ACTION AxisModules:
//*******************************************************************************************************************
// Moduli asse (Core: FB_AxisModule): ingressi dalla macchina, chiamate, uscite verso Safety e allarmi
//*******************************************************************************************************************
// In uso: per un asse aggiunto vale la presenza nei parametri macchina (Hmi.Param); per i sei assi storici le
// regole di prima. UR2 e UR_SIM: e' in uso uno solo dei due (ur2InUse); prima un'unica istanza di jog e di reset cambiava asse.
FOR i := 1 TO Mach.MAX_AXIS_CFG DO
	axisInUse[i] := Mach.aAxisCfg[i].bDefined AND Hmi.Param.aAxis[i].bPresent;
END_FOR
axisInUse[Mach.AX_USEL]		:= TRUE;
axisInUse[Mach.AX_USER]		:= TRUE;
axisInUse[Mach.AX_ERL]		:= TRUE;
axisInUse[Mach.AX_ERR]		:= TRUE;
axisInUse[Mach.AX_UR2]		:= ur2InUse;
axisInUse[Mach.AX_UR_SIM]	:= NOT ur2InUse;

// Ingressi comuni, dalla configurazione dell'asse (FB_MachineConfig)
mpgSelector := DINT_TO_UINT(stMpgEncoder.diSelector1);
FOR i := 1 TO Mach.MAX_AXIS_CFG DO
	IF Mach.aAxisCfg[i].bDefined THEN
		aAxisMod[i].bPowerEnable		:= axisInUse[i] AND motorsOn AND Safety.EmergenzaResettata;
		aAxisMod[i].fOverride			:= axisOverride;
		aAxisMod[i].bUseSoEReset		:= Mach.aAxisCfg[i].bSoEReset;
		aAxisMod[i].bSoEResetRequest	:= Safety.PulsanteResetEmergenza;
		aAxisMod[i].tPoweredOffDelay	:= tMotorsOffDelay;
		aAxisMod[i].bResetExecute		:= resetAxesCmd AND axisInUse[i];
		// Jog dal volantino: solo in manuale e con il ciclo fermo, l'asse scelto dal selettore.
		jogSelected := manualMode AND state = E_CycleState.Idle AND axisInUse[i]
			AND NOT calibStart[i] AND aAxisMod[i].nCalibrationStep = 0
			AND Mach.aAxisCfg[i].nMpgSelector <> 0 AND Mach.aAxisCfg[i].nMpgSelector = mpgSelector
			AND stMpgEncoder.diSafetySwitch;
		// Jog dall'HMI (stesse condizioni; i motori in manuale li tiene accesi il consenso del volantino).
		jogHmi := hmiConnected AND manualMode AND state = E_CycleState.Idle AND axisInUse[i] AND Hmi.Live.nJogAxis = i
			AND NOT calibStart[i] AND aAxisMod[i].nCalibrationStep = 0;
		aAxisMod[i].bJogForward			:= (jogSelected AND stMpgEncoder.eDirection = MC_Direction.MC_Positive_Direction)
			OR (jogHmi AND Hmi.Live.nJogDirection > 0);
		aAxisMod[i].bJogBackward		:= (jogSelected AND stMpgEncoder.eDirection = MC_Direction.MC_Negative_Direction)
			OR (jogHmi AND Hmi.Live.nJogDirection < 0);
		aAxisMod[i].fJogVelocity		:= Mach.aAxisCfg[i].fJogVelocity;
		aAxisMod[i].fJogAcceleration	:= Mach.aAxisCfg[i].fJogAcceleration;
		aAxisMod[i].fJogDeceleration	:= Mach.aAxisCfg[i].fJogDeceleration;
		aAxisMod[i].fJogJerk			:= Mach.aAxisCfg[i].fJogJerk;
		aAxisMod[i].bCalibrationStart	:= calibStart[i];
		aAxisMod[i].bUseCalibrationPos	:= calibUsePos[i];
		aAxisMod[i].fCalibrationPos		:= calibPos[i];
		aAxisMod[i].bWriteLimits		:= (i = limitsKickAxis);	// un asse alla volta (vedi fine AxisModules)
		// Limiti di un asse aggiunto dai parametri HMI; per gli assi storici li sovrascrive il blocco sotto.
		aAxisMod[i].fUpperLimit			:= Hmi.Param.aAxis[i].fUpperLimit;
		aAxisMod[i].fLowerLimit			:= Hmi.Param.aAxis[i].fLowerLimit;
	END_IF
END_FOR

// Calibrazione: comando e quota da HmiInputs (comando Calibrate), quota standard (GVL Calibration), datum di sicurezza
aAxisMod[Mach.AX_ERL].fHomePosition			:= Calibration.ERLHomePosition;
aAxisMod[Mach.AX_ERL].bDatumRequest			:= Safety.ERLDatumRequest;
aAxisMod[Mach.AX_ERL].bDatumDone			:= Safety.ERLDatumDone;

aAxisMod[Mach.AX_USEL].fHomePosition		:= Calibration.USELHomePosition;
aAxisMod[Mach.AX_USEL].bDatumRequest		:= Safety.USELDatumRquest;
aAxisMod[Mach.AX_USEL].bDatumDone			:= Safety.USELDatumDone;

aAxisMod[Mach.AX_UR2].fHomePosition			:= Calibration.URHomePosition;
aAxisMod[Mach.AX_UR2].bDatumRequest			:= Safety.URDatumRequest;
aAxisMod[Mach.AX_UR2].bDatumDone			:= Safety.URDatumDone;

aAxisMod[Mach.AX_ERR].fHomePosition			:= Calibration.ERRHomePosition;
aAxisMod[Mach.AX_ERR].bDatumRequest			:= Safety.ERRDatumRequest;
aAxisMod[Mach.AX_ERR].bDatumDone			:= Safety.ERRDatumDone;

aAxisMod[Mach.AX_USER].fHomePosition		:= Calibration.USERHomePosition;
aAxisMod[Mach.AX_USER].bDatumRequest		:= Safety.USERDatumRequest;
aAxisMod[Mach.AX_USER].bDatumDone			:= Safety.USERDatumDone;

// Limiti software dai parametri macchina (copia locale parametersRx). Il minimo delle USE non scende sotto
// il finecorsa della morsa montata (urUSE*MinPosition senza UR2, ur2USE*MinPosition con UR2).
aAxisMod[Mach.AX_ERL].fUpperLimit	:= parametersRx.ErLUpperLimit;
aAxisMod[Mach.AX_ERL].fLowerLimit	:= parametersRx.ErLLowerLimit;
aAxisMod[Mach.AX_USEL].fUpperLimit	:= parametersRx.UseLUpperLimit;
aAxisMod[Mach.AX_USEL].fLowerLimit	:= MAX(parametersRx.UseLLowerLimit, SEL(ur2InUse, urUSELMinPosition, ur2USELMinPosition));
aAxisMod[Mach.AX_UR2].fUpperLimit	:= parametersRx.UrRUpperLimit;
aAxisMod[Mach.AX_UR2].fLowerLimit	:= parametersRx.UrRLowerLimit;
aAxisMod[Mach.AX_ERR].fUpperLimit	:= parametersRx.ErRUpperLimit;
aAxisMod[Mach.AX_ERR].fLowerLimit	:= parametersRx.ErRLowerLimit;
aAxisMod[Mach.AX_USER].fUpperLimit	:= parametersRx.UseRUpperLimit;
aAxisMod[Mach.AX_USER].fLowerLimit	:= MAX(parametersRx.UseRLowerLimit, SEL(ur2InUse, urUSERMinPosition, ur2USERMinPosition));

// Chiamate (un asse NC per modulo)
aAxisMod[Mach.AX_USEL](stAxis := USEL);
aAxisMod[Mach.AX_USER](stAxis := USER);
aAxisMod[Mach.AX_ERL](stAxis := ERL);
aAxisMod[Mach.AX_ERR](stAxis := ERR);
aAxisMod[Mach.AX_UR2](stAxis := UR2);
aAxisMod[Mach.AX_UR_SIM](stAxis := UR_SIM);

// Uscite verso la sicurezza (lo stato della calibrazione per l'HMI e' in HmiOutputs)
// ERLDatumExecute non si azzera mai, come prima (la riga in InitCyclic era commentata): da verificare sullo schema safety.
IF aAxisMod[Mach.AX_ERL].bDatumExecute THEN
	Safety.ERLDatumExecute := TRUE;
END_IF
Safety.USELDatumExecute		:= aAxisMod[Mach.AX_USEL].bDatumExecute;
Safety.URDatumExecute		:= aAxisMod[Mach.AX_UR2].bDatumExecute;
Safety.ERRDatumExecute		:= aAxisMod[Mach.AX_ERR].bDatumExecute;
Safety.USERDatumExecute		:= aAxisMod[Mach.AX_USER].bDatumExecute;

// Esiti per la macchina a stati (letti nel ciclo dopo, come prima) e allarmi chiesti dai moduli
axesResetDone := TRUE;
axesResetError := FALSE;
axesResetErrorId := 0;
limitsBusy := FALSE;
FOR i := 1 TO Mach.MAX_AXIS_CFG DO
	IF Mach.aAxisCfg[i].bDefined THEN
		IF axisInUse[i] THEN
			axesResetDone := axesResetDone AND aAxisMod[i].bResetDone;
			IF aAxisMod[i].bResetError THEN
				axesResetError := TRUE;
				axesResetErrorId := MAX(axesResetErrorId, aAxisMod[i].nResetErrorId);
			END_IF
		END_IF
		limitsBusy := limitsBusy OR aAxisMod[i].bLimitsBusy;
		limitsFailed := limitsFailed OR aAxisMod[i].bLimitsError;
		CASE aAxisMod[i].eAlarm OF
			E_AxisAlarm.Calibration:
				RaiseAlarm(Id := Mach.aAxisCfg[i].nCalibrationAlarmId, Info := aAxisMod[i].nAlarmInfo);
			E_AxisAlarm.Limits:
				RaiseAlarm(Id := Mach.aAxisCfg[i].nLimitsAlarmId, Info := aAxisMod[i].nAlarmInfo);
		END_CASE
	END_IF
END_FOR

// Scrittura dei limiti un asse alla volta, come il vecchio ParameterWriteManager (MC_WriteParameter, non
// persistente: vedi FB_AxisModule). Un asse che fallisce non ferma i successivi.
// Fine: l'HMI aspetta Hmi.Sts.bWriteParametersDone FALSE -> TRUE (resta FALSE se un asse fallisce).
limitsKickAxis := 0;
IF limitsWriting AND NOT limitsBusy THEN
	FOR i := limitsAxis + 1 TO Mach.MAX_AXIS_CFG DO
		// asse simulato: nessun limite da scrivere
		IF limitsKickAxis = 0 AND Mach.aAxisCfg[i].bDefined AND i <> Mach.AX_UR_SIM THEN
			limitsKickAxis := i;
		END_IF
	END_FOR
	IF limitsKickAxis <> 0 THEN
		limitsAxis := limitsKickAxis;
	ELSE
		limitsWriting := FALSE;
		writeParametersDone := NOT limitsFailed;
	END_IF
END_IF
END_ACTION

ACTION DiagUpdate:
// Stato dei canali e storico dei cambi di passo nella GVL Diag (letta dall'HMI in un blocco).
FOR i := 0 TO 2 DO
	IF state = E_CycleState.HomingRun OR state = E_CycleState.HomingPrepare THEN
		Diag.Data.aChannel[i].bUsed := ProgramDB.homing.task[i].active;
	ELSE
		Diag.Data.aChannel[i].bUsed := ProgramDB.sequence[seqIdx].task[i].active;
	END_IF
	Diag.Data.aChannel[i].bDone := channelDone[i];
	Diag.Data.aChannel[i].bMWaiting := in_stNciToPlc[i].HskMFuncReq = 1 AND out_stPlcToNci[i].MFuncGranted = 0;
	IF in_stNciToPlc[i].HskMFuncReq = 1 THEN
		Diag.Data.aChannel[i].nMFunc := in_stNciToPlc[i].HskMFuncNo;
	ELSE
		Diag.Data.aChannel[i].nMFunc := 0;
	END_IF
	fbMFuncWait[i](IN := Diag.Data.aChannel[i].bMWaiting, PT := T#24H);
	Diag.Data.aChannel[i].tMWait := fbMFuncWait[i].ET;
	Diag.Data.aChannel[i].nItpState := udiItpState[i];
END_FOR
Diag.Data.aChannel[0].nLineNo := lineNo1;
Diag.Data.aChannel[1].nLineNo := lineNo2;
Diag.Data.aChannel[2].nLineNo := lineNo3;

// Sequenze attive: si ricontano solo quando arriva un programma nuovo (e al primo giro).
IF newProgramTrigger OR NOT diagSeqCounted THEN
	diagSeqCounted := TRUE;
	diagSeqIdx := 0;
	WHILE diagSeqIdx < Size.MAX_SEQUENCE AND_THEN ProgramDB.sequence[diagSeqIdx].active DO
		diagSeqIdx := diagSeqIdx + 1;
	END_WHILE
	Diag.Data.nSeqCount := diagSeqIdx;
END_IF

Diag.Data.eCycleEndReason := cycleEndReason;
IF state = E_CycleState.Centering THEN
	Diag.Data.nSubStep := fbCentering.nStep;
ELSE
	Diag.Data.nSubStep := fbSeq.eStep;
END_IF

fbDiagLog(
	nState		:= state,
	nSeqIdx		:= seqIdx,
	nAbortState	:= E_CycleState.Abort,
	nAlarmCount	:= Alarms.RaisedCount,
	nAlarmId	:= Alarms.LastRaisedId,
	nAlarmInfo	:= Alarms.LastRaisedInfo,
	stDiag		:= Diag.Data);
END_ACTION

ACTION DriveStatusManager:
// Calcola stato drive e consenso motori per HMI.
allDrivesEnabled := (bMotorsOnStatus[0] OR NOT Machine.parametersRx.USELPresent) AND 
					(bMotorsOnStatus[1] OR NOT Machine.parametersRx.ERLPresent) AND 
					(bMotorsOnStatus[2] OR NOT ur2InUse) AND 
					(bMotorsOnStatus[3] OR NOT Machine.parametersRx.USERPresent) AND
					(bMotorsOnStatus[4] OR NOT Machine.parametersRx.ERRPresent);
					
drivesError := (USEL.NcToPlc.ErrorCode <> 0 AND Machine.parametersRx.USELPresent) OR
			   (ERL.NcToPlc.ErrorCode <> 0 AND Machine.parametersRx.ERLPresent) OR
			   (USER.NcToPlc.ErrorCode <> 0 AND Machine.parametersRx.USERPresent) OR
			   (ERR.NcToPlc.ErrorCode <> 0 AND Machine.parametersRx.ERRPresent) OR
			   (UR2.NcToPlc.ErrorCode <> 0 AND ur2InUse);

//fbMotorsOffTrigger(CLK := allDrivesEnabled, Q => motorsOffTrigger);
fbSelectorOffTrigger(CLK := Safety.ModoAuto1Op, Q=> autoModeTrigger);

IF drivesError OR  motorsOffTrigger THEN
	motorsOn := FALSE;
END_IF
END_ACTION

ACTION HmiInputs:
//*******************************************************************************************************************
// Ingressi dall'HMI (GVL Hmi, contratto in docs/ADS_CONTRACT_V2.md) nelle variabili interne
//*******************************************************************************************************************
fbHmiWatchdog(nCounter := Hmi.Live.nWatchdog);
hmiConnected := fbHmiWatchdog.bAlive;

// Comandi con numero di sequenza: valgono un ciclo.
hmiStartCmd := FALSE;
hmiStopCmd := FALSE;
hmiResetCmd := FALSE;
hmiMotorsOnCmd := FALSE;
hmiMotorsOffCmd := FALSE;
hmiProgramLoadedCmd := FALSE;
hmiWriteParamsCmd := FALSE;
FOR i := 1 TO Mach.MAX_AXIS_CFG DO
	calibStart[i] := FALSE;
END_FOR

fbHmiCmd(stCmd := Hmi.Cmd);
IF fbHmiCmd.bNew THEN
	CASE Hmi.Cmd.eCommand OF
		E_HmiCommand.Start:
			hmiStartCmd := TRUE;
			fbHmiCmd.Ack(E_HmiResult.Accepted);
		E_HmiCommand.Stop:
			hmiStopCmd := TRUE;
			fbHmiCmd.Ack(E_HmiResult.Accepted);
		E_HmiCommand.Reset:
			hmiResetCmd := TRUE;
			fbHmiCmd.Ack(E_HmiResult.Accepted);
		E_HmiCommand.MotorsOn:
			hmiMotorsOnCmd := TRUE;
			fbHmiCmd.Ack(E_HmiResult.Accepted);
		E_HmiCommand.MotorsOff:
			hmiMotorsOffCmd := TRUE;
			fbHmiCmd.Ack(E_HmiResult.Accepted);
		E_HmiCommand.ProgramLoaded:
			hmiProgramLoadedCmd := TRUE;
			fbHmiCmd.Ack(E_HmiResult.Accepted);
		E_HmiCommand.WriteParameters:
			// Parametri macchina dell'HMI -> struttura persistente usata da tutto il PLC (Machine.parametersRx).
			Machine.parametersRx.EnableSirenOverride	:= Hmi.Param.bEnableSirenOverride;
			Machine.parametersRx.ERLPresent			:= Hmi.Param.aAxis[Mach.AX_ERL].bPresent;
			Machine.parametersRx.ERLCalibrated		:= Hmi.Param.aAxis[Mach.AX_ERL].bCalibrated;
			Machine.parametersRx.ERLCheckDone		:= Hmi.Param.aAxis[Mach.AX_ERL].bCheckDone;
			Machine.parametersRx.ErLUpperLimit		:= Hmi.Param.aAxis[Mach.AX_ERL].fUpperLimit;
			Machine.parametersRx.ErLLowerLimit		:= Hmi.Param.aAxis[Mach.AX_ERL].fLowerLimit;
			Machine.parametersRx.USELPresent		:= Hmi.Param.aAxis[Mach.AX_USEL].bPresent;
			Machine.parametersRx.USELCalibrated		:= Hmi.Param.aAxis[Mach.AX_USEL].bCalibrated;
			Machine.parametersRx.USELCheckDone		:= Hmi.Param.aAxis[Mach.AX_USEL].bCheckDone;
			Machine.parametersRx.UseLUpperLimit		:= Hmi.Param.aAxis[Mach.AX_USEL].fUpperLimit;
			Machine.parametersRx.UseLLowerLimit		:= Hmi.Param.aAxis[Mach.AX_USEL].fLowerLimit;
			Machine.parametersRx.UR2Present			:= Hmi.Param.aAxis[Mach.AX_UR2].bPresent;
			Machine.parametersRx.UR2Calibrated		:= Hmi.Param.aAxis[Mach.AX_UR2].bCalibrated;
			Machine.parametersRx.ER2CheckDone		:= Hmi.Param.aAxis[Mach.AX_UR2].bCheckDone;
			Machine.parametersRx.UrRUpperLimit		:= Hmi.Param.aAxis[Mach.AX_UR2].fUpperLimit;
			Machine.parametersRx.UrRLowerLimit		:= Hmi.Param.aAxis[Mach.AX_UR2].fLowerLimit;
			Machine.parametersRx.ERRPresent			:= Hmi.Param.aAxis[Mach.AX_ERR].bPresent;
			Machine.parametersRx.ERRCalibrated		:= Hmi.Param.aAxis[Mach.AX_ERR].bCalibrated;
			Machine.parametersRx.ERRCheckDone		:= Hmi.Param.aAxis[Mach.AX_ERR].bCheckDone;
			Machine.parametersRx.ErRUpperLimit		:= Hmi.Param.aAxis[Mach.AX_ERR].fUpperLimit;
			Machine.parametersRx.ErRLowerLimit		:= Hmi.Param.aAxis[Mach.AX_ERR].fLowerLimit;
			Machine.parametersRx.USERPresent		:= Hmi.Param.aAxis[Mach.AX_USER].bPresent;
			Machine.parametersRx.USERCalibrated		:= Hmi.Param.aAxis[Mach.AX_USER].bCalibrated;
			Machine.parametersRx.USERCheckDone		:= Hmi.Param.aAxis[Mach.AX_USER].bCheckDone;
			Machine.parametersRx.UseRUpperLimit		:= Hmi.Param.aAxis[Mach.AX_USER].fUpperLimit;
			Machine.parametersRx.UseRLowerLimit		:= Hmi.Param.aAxis[Mach.AX_USER].fLowerLimit;
			hmiWriteParamsCmd := TRUE;
			fbHmiCmd.Ack(E_HmiResult.Accepted);
		E_HmiCommand.Calibrate:
			IF Hmi.Cmd.nAxis < 1 OR Hmi.Cmd.nAxis > Mach.MAX_AXIS_CFG THEN
				fbHmiCmd.Ack(E_HmiResult.InvalidArgument);
			ELSIF NOT Mach.aAxisCfg[Hmi.Cmd.nAxis].bDefined OR Mach.aAxisCfg[Hmi.Cmd.nAxis].nCalibrationAlarmId = 0 THEN
				fbHmiCmd.Ack(E_HmiResult.InvalidArgument);		// asse senza calibrazione (es. UR_SIM)
			ELSIF NOT manualMode OR NOT Safety.ModoManuale OR state <> E_CycleState.Idle
				OR limitsWriting OR limitsRequest OR limitsStart OR aAxisMod[Hmi.Cmd.nAxis].bLimitsBusy THEN
				fbHmiCmd.Ack(E_HmiResult.Rejected);		// solo da fermo in manuale, senza scritture limiti
			ELSIF aAxisMod[Hmi.Cmd.nAxis].nCalibrationStep <> 0 THEN
				fbHmiCmd.Ack(E_HmiResult.Rejected);				// calibrazione gia' in corso
			ELSE
				calibStart[Hmi.Cmd.nAxis] := TRUE;
				calibUsePos[Hmi.Cmd.nAxis] := Hmi.Cmd.bFlag;
				calibPos[Hmi.Cmd.nAxis] := Hmi.Cmd.fValue;
				fbHmiCmd.Ack(E_HmiResult.Accepted);
			END_IF
		E_HmiCommand.SetCount:
			IF Hmi.Cmd.nValue >= 0 AND Hmi.Cmd.nValue <= 65535 THEN
				count := DINT_TO_UINT(Hmi.Cmd.nValue);
				fbHmiCmd.Ack(E_HmiResult.Accepted);
			ELSE
				fbHmiCmd.Ack(E_HmiResult.InvalidArgument);
			END_IF
	ELSE
		fbHmiCmd.Ack(E_HmiResult.UnknownCommand);
	END_CASE
END_IF

// Valori continui (Hmi.Live). Con l'HMI scollegata restano gli ultimi scritti, tranne il test uscite che si spegne.
hmiOverride := Hmi.Live.fOverride;
autoLoopMode := Hmi.Live.bLoopMode;
ncSingleBlock := Hmi.Live.nNcMode = 1;
hmiForce := hmiConnected AND Hmi.Live.bForceOutputs;
FOR i := 1 TO Mach.MAX_VALVE DO
	valveForce[i] := Hmi.Live.aValveForce[i];
END_FOR

// Pulsanti
hmiStop := hmiStopCmd;
hmiReset := hmiResetCmd;
END_ACTION

ACTION HmiOutputs:
//*******************************************************************************************************************
// Stato per l'HMI (GVL Hmi): configurazione e stato, un blocco ciascuno
//*******************************************************************************************************************
Hmi.Cfg.nInterfaceVersion	:= 2;
Hmi.Cfg.sMachine			:= 'Aut260045';
Hmi.Cfg.nMaxSequence		:= Size.MAX_SEQUENCE;
Hmi.Cfg.nMaxTask			:= Size.MAX_TASK;
Hmi.Cfg.nMaxAction			:= Size.MAX_ACTION;
Hmi.Cfg.nMaxPosition		:= Size.MAX_POSITION;
Hmi.Cfg.nMaxMacro			:= Size.MAX_MACRO;
Hmi.Cfg.nMaxAxisInGroup		:= Size.MAX_AXIS;
Hmi.Cfg.nChannels			:= Core_Param.MAX_CHANNEL;

FOR i := 1 TO Mach.MAX_AXIS_CFG DO
	Hmi.Cfg.aAxis[i].bDefined	:= Mach.aAxisCfg[i].bDefined;
	Hmi.Cfg.aAxis[i].sName		:= Mach.aAxisCfg[i].sName;
	Hmi.Cfg.aAxis[i].nOption	:= Mach.aAxisCfg[i].nMpgSelector;
	Hmi.Sts.aAxis[i].fActPos			:= Mach.aAxisCfg[i].fActPos;
	Hmi.Sts.aAxis[i].fActVelo			:= Mach.aAxisCfg[i].fActVelo;
	Hmi.Sts.aAxis[i].nErrorCode			:= Mach.aAxisCfg[i].nErrorCode;
	Hmi.Sts.aAxis[i].bEnabled			:= Mach.aAxisCfg[i].bDefined AND NOT Mach.aAxisCfg[i].bDisabled;
	Hmi.Sts.aAxis[i].bMoving			:= Mach.aAxisCfg[i].bMoving;
	Hmi.Sts.aAxis[i].bInUse				:= axisInUse[i];
	Hmi.Sts.aAxis[i].nCalibrationStep	:= aAxisMod[i].nCalibrationStep;
	Hmi.Sts.aAxis[i].bCalibrated		:= aAxisMod[i].bCalibrated;
	Hmi.Sts.aAxis[i].bLimitsBusy		:= aAxisMod[i].bLimitsBusy;
END_FOR
Hmi.Sts.aAxis[Mach.AX_ERL].fLastKnownPos	:= Machine.parametersTx.lastERLKnownPosition;
Hmi.Sts.aAxis[Mach.AX_USEL].fLastKnownPos	:= Machine.parametersTx.lastUSELKnownPosition;
Hmi.Sts.aAxis[Mach.AX_UR2].fLastKnownPos	:= Machine.parametersTx.lastUR2KnownPosition;
Hmi.Sts.aAxis[Mach.AX_ERR].fLastKnownPos	:= Machine.parametersTx.lastERRKnownPosition;
Hmi.Sts.aAxis[Mach.AX_USER].fLastKnownPos	:= Machine.parametersTx.lastUSERKnownPosition;

FOR i := 1 TO Mach.MAX_VALVE DO
	Hmi.Cfg.aValve[i].bDefined	:= Mach.aValve[i].pSet <> 0;
	Hmi.Cfg.aValve[i].sName		:= Mach.aValve[i].sName;
	Hmi.Cfg.aValve[i].nOption	:= SEL(Mach.aValve[i].eType = OUTPUT_ENUM.BISTABLE, 0, 1);
	IF Mach.aValve[i].pSet <> 0 THEN
		Hmi.Sts.aValve[i].bSet := Mach.aValve[i].pSet^;
	END_IF
	IF Mach.aValve[i].pReset <> 0 THEN
		Hmi.Sts.aValve[i].bReset := Mach.aValve[i].pReset^;
	END_IF
	IF Mach.aValve[i].pFbSet <> 0 THEN
		Hmi.Sts.aValve[i].bFbSet := Mach.aValve[i].pFbSet^;
	END_IF
	IF Mach.aValve[i].pFbReset <> 0 THEN
		Hmi.Sts.aValve[i].bFbReset := Mach.aValve[i].pFbReset^;
	END_IF
END_FOR

FOR i := 1 TO Core_Param.MAX_INPUT DO
	Hmi.Cfg.aInput[i].bDefined	:= Mach.aInput[i].pInput <> 0;
	Hmi.Cfg.aInput[i].sName		:= Mach.aInput[i].sName;
	IF Mach.aInput[i].pInput <> 0 THEN
		Hmi.Sts.aInput[i] := Mach.aInput[i].pInput^;
	END_IF
END_FOR

Hmi.Sts.nCmdAck				:= fbHmiCmd.nAck;
Hmi.Sts.eCmdResult			:= fbHmiCmd.eResult;
Hmi.Sts.bConnected			:= hmiConnected;
Hmi.Sts.nState				:= state;
Hmi.Sts.nSubStep			:= Diag.Data.nSubStep;
Hmi.Sts.eCycleEndReason		:= cycleEndReason;
Hmi.Sts.bIdle				:= programIdle;
Hmi.Sts.bCanExecute			:= programCanExecute;
Hmi.Sts.bRunning			:= programRunning;
Hmi.Sts.bStopped			:= programStopped;
Hmi.Sts.bAborted			:= programAborted;
Hmi.Sts.bHomingDone			:= homingDone;
Hmi.Sts.bManualMode			:= manualMode;
Hmi.Sts.bAutoMode			:= autoMode;
Hmi.Sts.bMotorsOn			:= allDrivesEnabled;
Hmi.Sts.bMotorsEnable		:= NOT drivesError;
Hmi.Sts.bLimitsWriting		:= limitsWriting;
Hmi.Sts.bWriteParametersDone := writeParametersDone;
Hmi.Sts.nCount				:= count;
Hmi.Sts.nSeqIdx				:= seqIdx;
Hmi.Sts.sProgramName		:= ProgramDB.parameters.prgName;
Hmi.Sts.aLineNo[0]			:= lineNo1;
Hmi.Sts.aLineNo[1]			:= lineNo2;
Hmi.Sts.aLineNo[2]			:= lineNo3;
FOR i := 0 TO 2 DO
	Hmi.Sts.aChannelDone[i] := channelDone[i];
END_FOR
Hmi.Sts.nMpgSelector		:= stMpgEncoder.diSelector1;
Hmi.Sts.nMpgSpeed			:= stMpgEncoder.diSelector2;
Hmi.Sts.aAlarmActive		:= Alarms.Active;
Hmi.Sts.aAlarmInfo			:= Alarms.Info;
END_ACTION

ACTION InitCyclic:
(*initialize data cyclic (every scan)*)
//*******************************************************************************************************************
// set FB defaults
//*******************************************************************************************************************
allDrivesEnabled	:= FALSE;
drivesError 		:= FALSE;


//Read Status
USEL.ReadStatus();
ERL.ReadStatus();
UR2.ReadStatus();
USER.ReadStatus();
ERR.ReadStatus();

resetAxesCmd								:= FALSE;	// FB_AxisModule: reset MC degli assi (passi 800 e 920)












fbMPGReadStatus.tUpdateTimerPt				:= T#5MS;
fbMPGReadStatus.uiScalingFactorDenominator	:= 300;
fbMPGReadStatus.uiScalingFactorNumerator	:= 1;
fbMpgReadStatus.uismoothingPercentage		:= 10;





parametersRx.ERLCalibrated					:= FALSE;
parametersRx.ERLPresent						:= FALSE;
parametersRx.ERRCalibrated					:= FALSE;
parametersRx.ERRPresent						:= FALSE;
parametersRx.UR2Calibrated					:= FALSE;
parametersRx.UR2Present						:= FALSE;
parametersRx.USELCalibrated					:= FALSE;
parametersRx.USELPresent					:= FALSE;
parametersRx.USERCalibrated					:= FALSE;
parametersRx.USERPresent					:= FALSE;
parametersRx.ERLCheckDone					:= FALSE;
parametersRx.USELCheckDone					:= FALSE;
parametersRx.ER2CheckDone					:= FALSE;
parametersRx.ERRCheckDone					:= FALSE;
parametersRx.USERCheckDone					:= FALSE;

fbCloseClampAfterCentering.IN				:= FALSE;
fbCloseClampAfterCentering.PT				:= T#1000MS;

waitForMove.IN 								:= FALSE;
waitForMove.PT 								:= T#1S;

startCondition								:= FALSE;
safeOverride								:= FALSE;
END_ACTION

ACTION InitOnce:
firstScan := FALSE;
END_ACTION

ACTION InputMapping:
//*******************************************************************************************************************
// Override, eventi dei comandi HMI, morsa in uso
//*******************************************************************************************************************
axisOverride 		:= hmiOverride;

IF ((USEL.NcToPlc.ActPos <= uselSafeOvPosition) AND USEL.Status.NegativeDirection) OR safety.ModoSemiAuto OR Safety.ModoManuale THEN
	IF hmiOverride > channel1SafeOverride THEN
		channel1Override := channel1SafeOverride;
	END_IF;
ELSE
	channel1Override := hmiOverride;
END_IF		

IF ((USER.NcToPlc.ActPos <= userSafeOvPosition) AND USER.Status.NegativeDirection) OR safety.ModoSemiAuto OR Safety.ModoManuale THEN
	IF hmiOverride > channel2SafeOverride THEN
		channel2Override := channel2SafeOverride;
	END_IF
ELSE
	channel2Override := hmiOverride;
END_IF		

IF (USER.NcToPlc.ActPos <= userSafeOvPosition AND USER.Status.NegativeDirection) OR (USEL.NcToPlc.ActPos <= uselSafeOvPosition AND USEL.Status.NegativeDirection) OR safety.ModoSemiAuto OR Safety.ModoManuale THEN
	IF hmiOverride > channel2SafeOverride	THEN
		channel3Override := channel2SafeOverride;
	END_IF
ELSE
	channel3Override := hmiOverride;
END_IF	


safeOverride := (USEL.NcToPlc.ActPos <= userSafeOvPosition AND USEL.Status.NegativeDirection) OR (USER.NcToPlc.ActPos <= userSafeOvPosition AND USER.Status.NegativeDirection);

IF hmiConnected THEN
	parametersRx := Machine.parametersRx;
END_IF

fbSelectorOnTrigger(CLK := Safety.ModoManuale, Q=> manualModeTrigger);
fbBimanualOpenClampTrigger(CLK := IO.bimanualOpenClamp, Q => bimanualOpenClampTriggerOut);

// Comandi dell'HMI (Hmi.Cmd): valgono un ciclo, come i fronti di prima.
startTriggerOut := hmiStartCmd;
writeParametersEvent := hmiWriteParamsCmd;

//*******************************************************************************************************************
// Nuovo programma dall'HMI (comando ProgramLoaded)
//*******************************************************************************************************************
newProgramTrigger := hmiProgramLoadedCmd;

//*******************************************************************************************************************
// Morsa per programma (ProgramDB.parameters.normalClamp)
//*******************************************************************************************************************
// Con la morsa normale il motore UR2 e' staccato: il programma usa l'asse simulato UR_SIM e
// non si controllano azionamento, allarme ed encoder dell'UR2. Il finecorsa minimo delle USE
// cambia (urUSE*MinPosition / ur2USE*MinPosition): quando la morsa cambia si riscrivono i limiti
// assi; la partenza ciclo aspetta la fine della scrittura (stato 0).
// UR2Present arriva solo con i parametri dell'HMI, quindi i limiti da riscrivere sono validi.
ur2InUse := Machine.parametersRx.UR2Present AND NOT ProgramDB.parameters.normalClamp;
IF writeParametersEvent THEN
	ur2InUsePrev := ur2InUse;
ELSIF ur2InUse <> ur2InUsePrev AND NOT limitsWriting THEN
	ur2InUsePrev := ur2InUse;
	limitsRequest := TRUE;
END_IF
END_ACTION

ACTION MacroManager:
//*******************************************************************************************************************
// Funzioni M dei canali NC
//*******************************************************************************************************************
// Cosa fa ogni funzione M (valvola, sincronismo, attesa, riga, start) e' scritto in una tabella in FB_MachineConfig;
// la esegue FB_MFuncDispatcher del Core. Qui restano solo le cose della macchina: interblocchi, flag di
// sincronismo storici, allarmi e abort chiesti dal dispatcher. La tabella la scrive fbMachineConfig (corpo di MAIN).

// Interblocchi: l'espulsore (M102) parte solo con l'UR2 entro 3 gradi da zero o con l'UR2 non usato.
Mach.aInterlock[Mach.IL_UR2_AT_ZERO] := ABS(UR2.NcToPlc.ActPos) < 3 OR NOT ur2InUse;

// Flag di sincronismo: le variabili storiche restano (azzeramenti nei passi del ciclo),
// il dispatcher lavora sui bit di syncFlags.
syncFlags := 0;
IF syncAck[0] THEN			syncFlags := syncFlags OR Mach.SYNC_ACK_L;		END_IF
IF syncAck[1] THEN			syncFlags := syncFlags OR Mach.SYNC_ACK_R;		END_IF
IF syncAck[2] THEN			syncFlags := syncFlags OR Mach.SYNC_ACK_UR2;	END_IF
IF UR2Done THEN				syncFlags := syncFlags OR Mach.SYNC_UR2_DONE;	END_IF
IF USEL_UR2_Ack THEN		syncFlags := syncFlags OR Mach.SYNC_UR2_ACK_L;	END_IF
IF USER_UR2_Ack THEN		syncFlags := syncFlags OR Mach.SYNC_UR2_ACK_R;	END_IF
IF USELDone THEN			syncFlags := syncFlags OR Mach.SYNC_DONE_L;		END_IF
IF USERDone THEN			syncFlags := syncFlags OR Mach.SYNC_DONE_R;		END_IF
IF UR2_USEL_Req THEN		syncFlags := syncFlags OR Mach.SYNC_UR2_REQ_L;	END_IF
IF UR2_USER_Req THEN		syncFlags := syncFlags OR Mach.SYNC_UR2_REQ_R;	END_IF

fbMFunc(
	bStart			:= startCondition,
	bCycleRunning	:= state > E_CycleState.Idle AND state < E_CycleState.Abort,
	nUnknownAlarmId	:= E_Alarm.UnknownMFunction,
	nDefCount		:= Mach.nMFuncCount,
	aNciToPlc		:= in_stNciToPlc,
	aPlcToNci		:= out_stPlcToNci,
	aDef			:= Mach.aMFunc,
	aValve			:= Mach.aValve,
	aInterlock		:= Mach.aInterlock,
	dwSyncFlags		:= syncFlags);

syncAck[0]		:= (syncFlags AND Mach.SYNC_ACK_L) <> 0;
syncAck[1]		:= (syncFlags AND Mach.SYNC_ACK_R) <> 0;
syncAck[2]		:= (syncFlags AND Mach.SYNC_ACK_UR2) <> 0;
UR2Done			:= (syncFlags AND Mach.SYNC_UR2_DONE) <> 0;
USEL_UR2_Ack	:= (syncFlags AND Mach.SYNC_UR2_ACK_L) <> 0;
USER_UR2_Ack	:= (syncFlags AND Mach.SYNC_UR2_ACK_R) <> 0;
USELDone		:= (syncFlags AND Mach.SYNC_DONE_L) <> 0;
USERDone		:= (syncFlags AND Mach.SYNC_DONE_R) <> 0;
UR2_USEL_Req	:= (syncFlags AND Mach.SYNC_UR2_REQ_L) <> 0;
UR2_USER_Req	:= (syncFlags AND Mach.SYNC_UR2_REQ_R) <> 0;

lineNo1 := fbMFunc.aLineNo[0];
lineNo2 := fbMFunc.aLineNo[1];
lineNo3 := fbMFunc.aLineNo[2];

// Allarmi e abort chiesti dal dispatcher: valvola senza conferma (Info = M), M sconosciuta (Info = canale*1000 + M).
FOR i:=0 TO 2 DO
	IF fbMFunc.aAlarmId[i] <> 0 THEN
		RaiseAlarm(Id := fbMFunc.aAlarmId[i], Info := fbMFunc.aAlarmInfo[i]);
	END_IF
END_FOR

IF fbMFunc.bAbort THEN
	state := E_CycleState.Abort;
END_IF

//*******************************************************************************************************************
// Time-out delle attese di sincronismo (M60, M61, M80, M110, M112, M113, M116) e dell'espulsione (M102)
//*******************************************************************************************************************
// Il manuale ferma la macchina con TIME OUT dopo circa 15 s di attesa (T51-T53). Qui il tempo conta solo
// mentre il ciclo non avanza: ogni canale e' finito, non e' usato dalla sequenza oppure aspetta una di queste
// funzioni. Un canale in movimento, una macro pneumatica (ha il suo time-out), un'attesa M130 o lo start del
// passo-passo (M95-M97) fermano il conteggio, cosi' un movimento lento non da' un falso time-out.
// Quali attese hanno il time-out e con quale allarme lo dice la tabella (nWaitAlarmId).
// Allo scadere: allarme con il numero della funzione M nel dettaglio e abort.
FOR i:=0 TO 2 DO
	syncWait[i] := fbMFunc.aWaiting[i];
	IF syncWait[i] THEN
		syncWaitAlarm[i] := fbMFunc.aWaitAlarmId[i];
	END_IF
END_FOR

// Solo con le tabelle in esecuzione: nel RUN la sequenza corrente, in INIT quella di posizionamento.
// In STOP (700-745) il conteggio si azzera e riparte da zero alla ripresa.
syncBlockedAll := state = E_CycleState.SeqRun OR state = E_CycleState.HomingRun;
FOR i:=0 TO 2 DO
	IF state = E_CycleState.HomingRun THEN
		syncTaskInUse := ProgramDB.homing.task[i].active;
	ELSE
		syncTaskInUse := ProgramDB.sequence[seqIdx].task[i].active;
	END_IF

	IF NOT (syncWait[i] OR channelDone[i] OR NOT syncTaskInUse) THEN
		syncBlockedAll := FALSE;
	END_IF
END_FOR

FOR i:=0 TO 2 DO
	fbSyncTimeOut[i](IN := syncWait[i] AND syncBlockedAll, PT := tSyncTimeOut);

	IF fbSyncTimeOut[i].Q THEN
		RaiseAlarm(Id := syncWaitAlarm[i], Info := in_stNciToPlc[i].HskMFuncNo);
		state := E_CycleState.Abort;
	END_IF
END_FOR
END_ACTION

ACTION Manual:
// Test uscite dall'HMI (HmiInputs): ogni valvola segue valveForce, la "reset" della bistabile e' il contrario.
IF hmiForce THEN
	FOR i := 1 TO Mach.MAX_VALVE DO
		IF Mach.aValve[i].pSet <> 0 THEN
			Mach.aValve[i].pSet^ := valveForce[i];
			IF Mach.aValve[i].pReset <> 0 THEN
				Mach.aValve[i].pReset^ := NOT valveForce[i];
			END_IF
		END_IF
	END_FOR
	// I bloccaggi pezzo 1 e 2 seguono i palpatori 1 e 2.
	IO.pc1centeringLock := valveForce[E_Valve.CenteringPiece1];
	IO.pc2centeringLock := valveForce[E_Valve.CenteringPiece2];
END_IF

IF state = E_CycleState.Idle THEN
	// Volantino: il selettore sceglie l'asse (ST_AxisCfg.nMpgSelector; il jog lo fa il suo FB_AxisModule, vedi
	// AxisModules) e le valvole dei pulsanti 1 e 3 (Mach.aMpgButton), che a ogni pressione si invertono.
	mpgSelector := DINT_TO_UINT(stMpgEncoder.diSelector1);
	mpgAxisSelected := FALSE;
	FOR i := 1 TO Mach.MAX_AXIS_CFG DO
		IF Mach.aAxisCfg[i].bDefined AND Mach.aAxisCfg[i].nMpgSelector <> 0 AND Mach.aAxisCfg[i].nMpgSelector = mpgSelector THEN
			mpgAxisSelected := TRUE;
		END_IF
	END_FOR

	IF mpgAxisSelected AND mpgSelector <= Mach.MAX_MPG_SEL THEN
		IF stMpgEncoder.uiSpeedDivider > 0 THEN
			axisOverride := LIMIT(
				0,
				stMpgEncoder.uiOverrideSpeed / stMpgEncoder.uiSpeedDivider,
				100
			);
		ELSE
			axisOverride := 0;
		END_IF;

		mpgValve := Mach.aMpgButton[mpgSelector, 1];
		IF stMpgEncoder.xButton1RTrigger AND mpgValve <> 0 THEN
			Mach.aValve[mpgValve].pSet^ := NOT Mach.aValve[mpgValve].pSet^;
			IF Mach.aValve[mpgValve].pReset <> 0 THEN
				Mach.aValve[mpgValve].pReset^ := NOT Mach.aValve[mpgValve].pSet^;
			END_IF
		END_IF

		mpgValve := Mach.aMpgButton[mpgSelector, 2];
		IF stMpgEncoder.xButton3RTrigger AND mpgValve <> 0 THEN
			Mach.aValve[mpgValve].pSet^ := NOT Mach.aValve[mpgValve].pSet^;
			IF Mach.aValve[mpgValve].pReset <> 0 THEN
				Mach.aValve[mpgValve].pReset^ := NOT Mach.aValve[mpgValve].pSet^;
			END_IF
		END_IF
	END_IF
ELSE
	IF state = E_CycleState.SeqRun THEN
		IF stMpgEncoder.uiSpeedDivider > 0 THEN
			channel1Override := LIMIT(0,stMpgEncoder.uiOverrideSpeed/stMpgEncoder.uiSpeedDivider,channel1SafeOverride);
			channel2Override := LIMIT(0,stMpgEncoder.uiOverrideSpeed/stMpgEncoder.uiSpeedDivider,channel2SafeOverride);
			channel3Override := LIMIT(0,stMpgEncoder.uiOverrideSpeed/stMpgEncoder.uiSpeedDivider,channel3SafeOverride);
		ELSE
			channel1Override := 0;
			channel2Override := 0;
			channel3Override := 0;
		END_IF
	END_IF
	
	IF state = E_CycleState.Centering THEN
		IF stMpgEncoder.uiSpeedDivider > 0 THEN
			axisOverride := LIMIT(0,stMpgEncoder.uiOverrideSpeed/stMpgEncoder.uiSpeedDivider,channel1SafeOverride);
		ELSE
			axisOverride := 0;
		END_IF
	END_IF
END_IF



// Calibrazioni degli assi: in FB_AxisModule (action AxisModules).
END_ACTION

ACTION MotorStatusManager:
// Aggiorna richiesta motori e stato manuale.
fbTimerOffMotos[0](IN := NOT USEL.Status.Disabled, PT := tMotorsOffDelay, Q=> bMotorsOnStatus[0]);
fbTimerOffMotos[1](IN := NOT ERL.Status.Disabled, PT := tMotorsOffDelay, Q=> bMotorsOnStatus[1]);
fbTimerOffMotos[2](IN := NOT UR2.Status.Disabled, PT := tMotorsOffDelay, Q=> bMotorsOnStatus[2]);
fbTimerOffMotos[3](IN := NOT USER.Status.Disabled, PT := tMotorsOffDelay, Q=> bMotorsOnStatus[3]);
fbTimerOffMotos[4](IN := NOT ERR.Status.Disabled, PT := tMotorsOffDelay, Q=> bMotorsOnStatus[4]);

IF hmiMotorsOnCmd THEN
	motorsOn := TRUE;
END_IF
IF hmiMotorsOffCmd THEN
	motorsOn := FALSE;
END_IF

IF manualMode THEN
	motorsOn := stMpgEncoder.diSafetySwitch; 
END_IF
END_ACTION

ACTION OutputMapping:
//*******************************************************************************************************************
// Mapping digital outputs  
//*******************************************************************************************************************

IO.smc1[0].0 := IO.erLeftOutReset;
IO.smc1[0].1 := IO.erLeftOutSet;
IO.smc1[0].2 := IO.erRightOutReset;
IO.smc1[0].3 := IO.erRightOutSet;
IO.smc1[0].4 := IO.useLeftUpReset;
IO.smc1[0].5 := IO.useLeftUpSet;
IO.smc1[0].6 := IO.useRightUpReset;
IO.smc1[0].7 := IO.useRightUpSet;

IO.smc1[1].0 := IO.epLeftOutSet;
IO.smc1[1].1 := IO.epLeftOutReset;
IO.smc1[1].2 := IO.epLeftBend;
IO.smc1[1].3 := NOT IO.epLeftBend;
IO.smc1[1].4 := IO.epRightOutSet;
IO.smc1[1].5 := IO.epRightOutReset;
IO.smc1[1].6 := IO.epRightBend;
IO.smc1[1].7 := NOT IO.epRightBend;

IO.smc1[2].0 := IO.supportLeftOutSet;
IO.smc1[2].1 := IO.supportLeftOutReset;
IO.smc1[2].2 := IO.supportRightOutSet;
IO.smc1[2].3 := IO.supportRightOutReset;
IO.smc1[2].4 := IO.clampClosedSet;
IO.smc1[2].5 := IO.clampClosedReset;
IO.smc1[2].6 := IO.clampEjectSet;
IO.smc1[2].7 := IO.clampEjectReset;


IO.smc2[0].0 := IO.centringClamp1Left;
IO.smc2[0].2 := IO.centringClamp2Left;
IO.smc2[0].4 := IO.centringClamp3Left;
IO.smc2[0].6 := IO.centringClamp4Left;
IO.smc2[1].0 :=  IO.centeringLeft1Set;
IO.smc2[1].2 :=  IO.centeringLeft2Set;
IO.smc2[1].4 :=  IO.centeringLeft3Set;
IO.smc2[1].6 :=  IO.centeringLeft4Set;

IO.smc2[2].0 := IO.centeringLeftReset;
IO.smc2[2].2 := IO.centringSet;
IO.smc2[2].3 := IO.centringReset;
IO.smc2[2].4 := IO.centringClampSet;
io.smc2[2].6 := io.centeringOutSet;


IO.chillerEnabled := TRUE;

stTwoHandControl.doStartLED := (programCanExecute AND NOT programRunning) OR (programRunning AND Clock.pulse2Hz);
stTwoHandControl.doStopLED	:= programRunning;

IO.turretGreen := programRunning;
IO.spiaPulsanteStop := programRunning;

// Spia start: in automatico, a macchina ferma e senza allarmi bloccanti.
IO.spiaPulsanteStart := autoMode AND NOT programRunning AND Alarms.CountBlocking = 0;

IO.turretYellow := manualMode OR (autoMode AND Clock.pulse2Hz AND NOT programRunning);
IO.turretRed := Alarms.CountBlocking > 0;

IO.turretSiren := (safeOverride AND (Clock.pulse2Hz) AND programRunning) AND parametersRx.EnableSirenOverride;

//IF autoMode THEN
//	IO.turretSiren := (safeOverride AND (Clock.pulse2Hz) AND programRunning) AND parametersRx.EnableSirenOverride;
//ELSE
//	IO.turretSiren := (safeOverride AND (Clock.pulse2Hz)) AND parametersRx.EnableSirenOverride;
//END_IF

IF parametersRx.ERLCalibrated AND parametersRx.ERLCheckDone THEN
	Machine.parametersTx.lastERLKnownPosition := ERL.NcToPlc.ActPos;
END_IF

IF parametersRx.USELCalibrated AND parametersRx.USELCheckDone THEN
	Machine.parametersTx.lastUSELKnownPosition := USEL.NcToPlc.ActPos;
END_IF

// Con la morsa normale l'encoder UR2 e' staccato: non si sovrascrive l'ultima posizione buona.
IF parametersRx.UR2Calibrated AND parametersRx.ER2CheckDone AND ur2InUse THEN
	Machine.parametersTx.lastUR2KnownPosition := UR2.NcToPlc.ActPos;
END_IF

IF parametersRx.ERRCalibrated AND parametersRx.ERRCheckDone THEN
	Machine.parametersTx.lastERRKnownPosition := ERR.NcToPlc.ActPos;
END_IF

IF parametersRx.USERCalibrated AND parametersRx.USERCheckDone THEN
	Machine.parametersTx.lastUSERKnownPosition := USER.NcToPlc.ActPos;
END_IF
END_ACTION

ACTION ParameterWriteManager:
// Scrittura dei limiti software degli assi: su comando dell'HMI (WriteParameters) o quando cambia la morsa
// (limitsRequest, InputMapping). Ogni FB_AxisModule scrive massimo e minimo del suo asse; AxisModules
// li avvia un asse alla volta e valuta la fine. Mentre si scrive la partenza ciclo aspetta (passo 0).
limitsStart := writeParametersEvent OR limitsRequest;
limitsRequest := FALSE;

IF limitsStart THEN
	// L'HMI aspetta Done FALSE -> TRUE per ogni scrittura.
	writeParametersDone := FALSE;
	limitsWriting := TRUE;
	limitsFailed := FALSE;
	limitsAxis := 0;		// si riparte dal primo asse (AxisModules)
END_IF
END_ACTION

ACTION SafetyManager:
//*******************************************************************************************************************
// Sefety
//*******************************************************************************************************************

IF (Safety.ComErr OR Safety.FBErr OR Safety.OtherErr) THEN
	Safety.Run := Clock.pulse5Hz;
	Safety.Ack := Safety.PulsanteResetEmergenza;
ELSE
	Safety.Run := TRUE;
	Safety.Ack := FALSE;
END_IF

IF (Safety.USEL_ERL_ComErr OR Safety.USEL_ERL_FBErr OR Safety.USEL_ERL_OtherErr) THEN
	Safety.USEL_ERL_Run := Clock.pulse5Hz;
	Safety.USEL_ERL_Ack := Safety.PulsanteResetEmergenza;
ELSE
	Safety.USEL_ERL_Run := TRUE;
	Safety.USEL_ERL_Ack := FALSE;
END_IF

IF (Safety.USER_ERR_ComErr OR Safety.USER_ERR_FBErr OR Safety.USER_ERR_OtherErr) THEN
	Safety.USER_ERR_Run := Clock.pulse5Hz;
	Safety.USER_ERR_Ack := Safety.PulsanteResetEmergenza;
ELSE
	Safety.USER_ERR_Run := TRUE;
	Safety.USER_ERR_Ack := FALSE;
END_IF

IF (Safety.UR_ComErr OR Safety.UR_FBErr OR Safety.UR_OtherErr) THEN
	Safety.UR_Run := Clock.pulse5Hz;
	Safety.UR_Ack := Safety.PulsanteResetEmergenza;
ELSE
	Safety.UR_Run := TRUE;
	Safety.UR_Ack := FALSE;
END_IF

Safety.ResetEmergenza := safety.PulsanteResetEmergenza;
Safety.ResetBarriere := safety.PulsanteResetBarriere; 
Safety.ERLCommErrorAck :=  Safety.PulsanteResetEmergenza;
Safety.USELCommErrorAck	:=  Safety.PulsanteResetEmergenza;
Safety.URCommErrorAck :=  Safety.PulsanteResetEmergenza;
Safety.ERRCommErrorAck :=  Safety.PulsanteResetEmergenza;
Safety.USERCommErrorAck :=  Safety.PulsanteResetEmergenza;

IF  Safety.PulsanteResetEmergenza  THEN
	Safety.Ack := TRUE;
	Safety.ERLSafetyReset := 1;
	Safety.USELSafetyReset := 1;
	Safety.URSafetyReset := 1;
	Safety.ERRSafetyReset := 1;
	Safety.USERSafetyReset := 1;
ELSE
	Safety.ERLSafetyReset := 0;
	Safety.USELSafetyReset := 0;
	Safety.URSafetyReset := 0;
	Safety.ERRSafetyReset := 0;
	Safety.USERSafetyReset := 0;
END_IF

Safety.SpiaPulsanteRipristinoSicurezze := (NOT Safety.EmergenzaResettata AND Clock.pulse2Hz) OR Safety.EmergenzaResettata;
Safety.SpiaPulsanteRipristinoBarriere := (NOT Safety.BarriereResettate AND Clock.pulse2Hz) OR Safety.BarriereResettate;
END_ACTION

ACTION StateMachine:
//*******************************************************************************************************************
// State machine
//*******************************************************************************************************************
IF manualMode THEN
	IF stMpgEncoder.xbutton2RTrigger THEN
		startCondition := TRUE;
	END_IF
ELSIF autoMode THEN
	IF startTriggerOut OR stTwoHandControl.xStartRTrigger OR stTwoHandControl.xTwoHandRTrigger THEN
		startCondition := TRUE;
	END_IF
END_IF

//*******************************************************************************************************************
// Blocca lo start anche se calibrazione e pulsante Start arrivano nella stessa scansione.
// I comandi calibStart sono gia' acquisiti da HmiInputs; gli esiti dei moduli sono del ciclo precedente.
//*******************************************************************************************************************
calibrationBusy := FALSE;
FOR i := 1 TO Mach.MAX_AXIS_CFG DO
	calibrationBusy := calibrationBusy OR calibStart[i] OR aAxisMod[i].nCalibrationStep <> 0;
END_FOR

//*******************************************************************************************************************
// Gruppi e tabelle NC della sequenza (Core: FB_SequenceRunner)
//*******************************************************************************************************************
// Il comando viene dal passo del ciclo; il runner gira prima del CASE, cosi' i passi leggono il suo esito
// nello stesso ciclo (come prima, quando le tabelle si chiamavano dentro i passi). Va chiamato sempre:
// con None fa solo girare i FB dei gruppi.
CASE state OF
	E_CycleState.SeqPrepare, E_CycleState.HomingPrepare:
		seqCmd := E_SeqCmd.Prepare;
	E_CycleState.SeqRun, E_CycleState.HomingRun:
		seqCmd := E_SeqCmd.Run;
	E_CycleState.ResumeResetTables, E_CycleState.ResumeResetWait:
		seqCmd := E_SeqCmd.ResetTables;
ELSE
	seqCmd := E_SeqCmd.None;
END_CASE

IF state = E_CycleState.HomingPrepare OR state = E_CycleState.HomingRun THEN
	fbSeq.pSequence := ADR(ProgramDB.homing);
ELSE
	fbSeq.pSequence := ADR(ProgramDB.sequence[seqIdx]);
END_IF

fbSeq(
	eCmd					:= seqCmd,
	nGroupIdBase			:= Mach.NC_GROUP_BASE,
	bCenteringCorrection	:= ProgramDB.parameters.centering >= CENTERING_ENUM.TB,
	fToleranceMeasure		:= ToleranceMeasure,
	bSingleBlock			:= ncSingleBlock,
	nDefCount				:= Mach.nMFuncCount,
	bLogFeederEntries		:= bLogEntries[0],
	aNciToPlc				:= in_stNciToPlc,
	aAxisCfg				:= Mach.aAxisCfg,
	aDef					:= Mach.aMFunc);

// Centraggio TL/TB (FB della macchina): chiamato sempre, perche' FB di movimento e timer girino a ogni ciclo.
fbCentering(
	bExecute		:= state = E_CycleState.Centering,
	bStart			:= startCondition,
	bStepMode		:= ncSingleBlock,
	fMoveSpeed		:= USEMoveSpeed,
	fSearchSpeed	:= USESearchSpeed,
	nGroupIdBase	:= Mach.NC_GROUP_BASE,
	stUseL			:= USEL,
	stUseR			:= USER);

// Arresto, step-on e reset dei canali NC (Core: FB_NcChannels): il comando viene dal passo del ciclo,
// i passi leggono bDone/bError nello stesso ciclo.
CASE state OF
	E_CycleState.Abort, E_CycleState.Stop, E_CycleState.ToManualEStop:
		ncCmd := E_NcChannelCmd.EStop;
	E_CycleState.Resume:
		IF lastState = E_CycleState.SeqRun THEN
			ncCmd := E_NcChannelCmd.StepOn;
		ELSE
			ncCmd := E_NcChannelCmd.None;
		END_IF
	E_CycleState.ResetChannels:
		ncCmd := E_NcChannelCmd.Reset;
ELSE
	ncCmd := E_NcChannelCmd.None;
END_CASE

fbNc(eCmd := ncCmd, aNciToPlc := in_stNciToPlc);

CASE state OF
	(*********************** IDLE **********************)
	E_CycleState.Idle:	
		// Con una scrittura limiti assi in corso (es. cambio morsa) la partenza aspetta.
		IF startCondition AND NOT limitsWriting AND NOT calibrationBusy THEN
			state := E_CycleState.StartChecks;
		END_IF
		
		IF hmiReset THEN
			state := E_CycleState.Reset;
		END_IF
		
		IF stTwoHandControl.xStopButtonDelayTrigger THEN
			IO.clampClosedReset := TRUE;
			IO.clampClosedSet 	:= FALSE;
		END_IF

		// L'operatore ha azzerato o corretto il contapezzi dall'HMI (comando SetCount): l'avviso si spegne.
		IF Alarms.Active[E_Alarm.BatchCompleted]
			AND NOT (ProgramDB.parameters.pcsCounter > 0 AND count >= ProgramDB.parameters.pcsCounter) THEN
			Alarms.Active[E_Alarm.BatchCompleted] := FALSE;
		END_IF

	E_CycleState.StartChecks:
		state := E_CycleState.SeqInit;

		// I messaggi "start rifiutato" valgono per l'ultimo tentativo.
		Alarms.Active[E_Alarm.StartDriveError]		:= FALSE;
		Alarms.Active[E_Alarm.StartMotorsOff]		:= FALSE;
		Alarms.Active[E_Alarm.StartNoProgram]		:= FALSE;
		Alarms.Active[E_Alarm.StartCabinetAlarm]	:= FALSE;
		Alarms.Active[E_Alarm.BatchCompleted]		:= FALSE;

		// Lotto completato: niente start finche' l'operatore non azzera o corregge il contapezzi.
		// pcsCounter = 0: nessun lotto.
		IF ProgramDB.parameters.pcsCounter > 0 AND count >= ProgramDB.parameters.pcsCounter THEN
			RaiseAlarm(Id := E_Alarm.BatchCompleted);
			state := E_CycleState.Idle;
		END_IF

		IF Alarms.StartBlockedByCabinet THEN
			RaiseAlarm(Id := E_Alarm.StartCabinetAlarm);
			state := E_CycleState.Idle;
		END_IF

		IF drivesError THEN 
			RaiseAlarm(Id := E_Alarm.StartDriveError);
			state := E_CycleState.Idle;
		END_IF
		
		IF NOT allDrivesEnabled THEN 
			RaiseAlarm(Id := E_Alarm.StartMotorsOff);
			state := E_CycleState.Idle;
		END_IF
		
		IF NOT ProgramDB.sequence[0].active THEN
			RaiseAlarm(Id := E_Alarm.StartNoProgram);
			state := E_CycleState.Idle;
		END_IF

		IF state = E_CycleState.Idle THEN
			cycleEndReason := E_CycleEndReason.StartRefused;
		ELSE
			cycleEndReason := E_CycleEndReason.None;
		END_IF

	(*********************** CENTERING **********************)
	E_CycleState.CenteringSelect:	 
		IF homingDone THEN
			CASE ProgramDB.parameters.centering OF
				CENTERING_ENUM.NO:	//Esclusione Centratore.
					state := E_CycleState.SeqInit;
				
				CENTERING_ENUM.TL:	//Centratore predisposto per la ripresa della tolleranza nei terminali del pezzo.	
					state := E_CycleState.Centering;

				CENTERING_ENUM.TB:	//Centratore predisposto per la ripresa della tolleranza in un curva (tutta la tolleranza in una curva) oppure in due curve (metà tolleranza in una curva, metà tolleranza in un'altra curva) oppure in tre o quattro curve.
					state := E_CycleState.Centering;
			ELSE
				// ACC (centraggio automatico) o valore sconosciuto: non implementato, prima la macchina restava ferma qui.
				RaiseAlarm(Id := E_Alarm.CenteringModeNotSupported, Info := TO_UDINT(ProgramDB.parameters.centering));
				state := E_CycleState.Abort;
			END_CASE
		ELSE
			state := E_CycleState.HomingPrepare;
		END_IF

	(*********************** Centraggio TL/TB (FB_Centering) **********************)
	// Le fasi (ex passi 55-78) sono in fbCentering, chiamato in testa con bExecute in questo passo;
	// il passo interno e' in Diag.Data.nSubStep. Qui restano solo le uscite verso il ciclo.
	E_CycleState.Centering:

		IF fbCentering.bDone THEN
			IF ProgramDB.parameters.centering = CENTERING_ENUM.TB THEN
				MeasureL := fbCentering.fMeasureL;
				MeasureR := fbCentering.fMeasureR;
				ToleranceMeasure := MeasureL + MeasureR;
			END_IF

			// Fine del centraggio: uno stop premuto durante la fase si applica qui, la ripresa va alla prima riga.
			IF stopPending THEN
				lastState := E_CycleState.SeqInit;
				state := E_CycleState.Stop;
			ELSE
				state := E_CycleState.SeqInit;
			END_IF

		ELSIF fbCentering.bFailed THEN
			// Pezzo gia' presente o non trovato (allarmi 61/62): si rifa' il posizionamento iniziale.
			homingDone := FALSE;
			IF stopPending THEN
				lastState := E_CycleState.HomingPrepare;
				state := E_CycleState.Stop;
			ELSE
				state := E_CycleState.HomingPrepare;
			END_IF

		ELSIF fbCentering.bAbort THEN
			// Errore NC (allarmi 200-205, gia' memorizzati da fbCentering).
			state := E_CycleState.Abort;
		END_IF

	(*********************** INIT Before execution **********************)  
	E_CycleState.SeqInit:	
		//PrintProgram();
		seqIdx := 0;
		
		USELDone := FALSE;
		USERDone := FALSE;
		UR2Done	:= FALSE;
		USEL_UR2_Ack := FALSE;
		USER_UR2_Ack := FALSE;
		UR2_USEL_Req := FALSE;
		UR2_USER_Req := FALSE;
		
		IF homingDone THEN
			state := E_CycleState.SeqPrepare;
		ELSE
			state := E_CycleState.HomingPrepare;
		END_IF
	
	(*********************** Preparazione della sequenza **********************)
	// Reset e costruzione dei gruppi NC, tabelle, invio ai canali: fbSeq (FB_SequenceRunner) con il comando
	// Prepare dato in testa alla macchina a stati. Gli allarmi restano quelli dei vecchi passi 120-400.
	E_CycleState.SeqPrepare:
		IF fbSeq.bReady THEN
			// Un canale senza task in questa sequenza e' gia' finito: altrimenti lo stato 410 lo aspetterebbe per sempre.
			FOR i:=0 TO 2 DO
				channelDone[i] := NOT ProgramDB.sequence[seqIdx].task[i].active;
			END_FOR
			state := E_CycleState.SeqRun;
		END_IF

		IF fbSeq.bError THEN
			CASE fbSeq.eErrorStep OF
				E_SeqStep.ClearGroups:	seqAlarmId := E_Alarm.NcClearGroups;
				E_SeqStep.BuildGroups:	seqAlarmId := E_Alarm.NcBuildGroups;
				E_SeqStep.TableReset:	seqAlarmId := E_Alarm.NcFeedTableReset;
				E_SeqStep.TableFeed:	seqAlarmId := E_Alarm.NcFeedTableStart;
			ELSE
				seqAlarmId := E_Alarm.NcFeedTablePrep;
			END_CASE
			RaiseAlarm(Id := seqAlarmId, Info := fbSeq.nErrorId);
			state := E_CycleState.Abort;
		END_IF

	(*********************** Preparazione dell'homing (posizionamento iniziale) **********************)
	E_CycleState.HomingPrepare:
		IO.centringSet := FALSE;
		IO.centringReset := TRUE;
		IO.centringLeftUpSet := FALSE;
		IO.centringLeftUpReset := TRUE;
		IO.centringRightUpSet := FALSE;
		IO.centringRightUpReset := TRUE;
		IO.centringClamp1Left := FALSE;
		IO.centringClamp2Left := FALSE;
		IO.centringClamp3Left := FALSE;
		IO.centringClamp4Left := FALSE;
		IO.centeringLeft1Set := FALSE;
		IO.centeringLeft2Set := FALSE;
		IO.centeringLeft3Set := FALSE;
		IO.centeringLeft4Set := FALSE;
		IO.centringClampSet := FALSE;

		IF fbSeq.bReady THEN
			// Come per le sequenze: un canale senza task nell'homing e' gia' finito.
			FOR i:=0 TO 2 DO
				channelDone[i] := NOT ProgramDB.homing.task[i].active;
				syncAck[i] := FALSE;
			END_FOR
			state := E_CycleState.HomingRun;
		END_IF

		IF fbSeq.bError THEN
			CASE fbSeq.eErrorStep OF
				E_SeqStep.ClearGroups:	seqAlarmId := E_Alarm.NcClearGroupsInit;
				E_SeqStep.BuildGroups:	seqAlarmId := E_Alarm.NcBuildGroupsInit;
				E_SeqStep.TableReset:	seqAlarmId := E_Alarm.NcFeedTableResetInit;
				E_SeqStep.TableFeed:	seqAlarmId := E_Alarm.NcFeedTableStartInit;
			ELSE
				seqAlarmId := E_Alarm.NcFeedTablePrepInit;
			END_CASE
			RaiseAlarm(Id := seqAlarmId, Info := fbSeq.nErrorId);
			state := E_CycleState.Abort;
		END_IF

	(*********************** Run **********************)  
	E_CycleState.SeqRun:	
		
		// Fine dei canali dal runner (comando Run): si memorizza qui.
		FOR i:=0 TO 2 DO
			IF fbSeq.aChannelDone[i] THEN
				channelDone[i] := TRUE;
			END_IF
		END_FOR

		// Fine sequenza: ogni ramo lascia lo stato 410 nella stessa scansione, cosi' la fine pezzo
		// (contapezzi, lotto) si valuta una volta sola anche se channelDone[] restano TRUE.
		IF channelDone[0] AND channelDone[1] AND channelDone[2] THEN
			homingDone := FALSE;

			IF seqIdx < Size.MAX_SEQUENCE - 1 THEN
				nextSequenceActive := ProgramDB.sequence[seqIdx + 1].active;
			ELSE
				nextSequenceActive := FALSE;
			END_IF

			IF nextSequenceActive THEN
				seqIdx := seqIdx + 1;
				State := E_CycleState.SeqPrepare;
			ELSE
				// Fine pezzo. Il contapezzi sale sempre (senza superare il massimo di UINT);
				// con pcsCounter > 0 il lotto completato ferma la macchina, qualunque sia il modo di espulsione.
				seqIdx := 0;
				count := UDINT_TO_UINT(MIN(count + ProgramDB.parameters.pcsCycle, UDINT#65535));

				IF ProgramDB.parameters.pcsCounter > 0 AND count >= ProgramDB.parameters.pcsCounter THEN
					RaiseAlarm(Id := E_Alarm.BatchCompleted);
					cycleEndReason := E_CycleEndReason.BatchCompleted;
					State := E_CycleState.CycleEnd;
				ELSIF newProgramPending THEN
					// Nuovo programma caricato dall'HMI: il ciclo si chiude qui invece di
					// ripartire con i dati vecchi. Il reset viene applicato in stato 850.
					cycleEndReason := E_CycleEndReason.NewProgram;
					State := E_CycleState.CycleEnd;
				ELSIF autoLoopMode THEN
					cycleEndReason := E_CycleEndReason.PieceDone;
					CASE ProgramDB.parameters.ejectMode OF
						EJECT_ENUM.YES:
							state := E_CycleState.CenteringSelect;

						EJECT_ENUM.NO_2_START:
							state := E_CycleState.WaitStartNextPiece;

						EJECT_ENUM.NO_1_START:
							state := E_CycleState.CenteringSelect;
					ELSE
						// modo sconosciuto (es. il vecchio EJECT 3): fine ciclo
						cycleEndReason := E_CycleEndReason.UnknownEjectMode;
						State := E_CycleState.CycleEnd;
					END_CASE
				ELSE
					cycleEndReason := E_CycleEndReason.SingleCycle;
					State := E_CycleState.CycleEnd;
				END_IF
			END_IF
		END_IF
		
		IF fbSeq.bError THEN
			RaiseAlarm(Id := E_Alarm.NcFeedTableRun, Info := fbSeq.nErrorId);
			state := E_CycleState.Abort;
		END_IF
	
	(*********************** Run Init **********************)  
	E_CycleState.HomingRun:	
		IO.centeringLeftReset := TRUE;
		IO.centeringRightReset := TRUE;
		
		FOR i:=0 TO 2 DO
			IF fbSeq.aChannelDone[i] THEN
				channelDone[i] := TRUE;
			END_IF
		END_FOR

		IF channelDone[0] AND channelDone[1] AND channelDone[2]  THEN 
			homingDone := TRUE;
			
			IF ProgramDB.parameters.centering <> CENTERING_ENUM.NO THEN
				IO.centeringLeft1Set := TRUE;
				IO.centeringLeft2Set := TRUE;
				IO.centeringLeft3Set := TRUE;
				IO.centeringLeft4Set := TRUE;
				IO.centringSet := TRUE;
				IO.centringReset := FALSE;
				IO.centringClamp1Left := FALSE;
				IO.centringClamp2Left := FALSE;
				IO.centringClamp3Left := FALSE;
				IO.centringClamp4Left := FALSE;
				IO.centringClampSet := FALSE;
			END_IF

			// Fine del posizionamento iniziale: uno stop premuto durante la fase (o durante l'attesa
			// dello start) si applica qui; lo start della ripresa fa partire il centraggio (stato 50).
			IF stopPending THEN
				lastState := E_CycleState.CenteringSelect;
				state := E_CycleState.Stop;
			ELSIF startCondition THEN
				state := E_CycleState.CenteringSelect;
			END_IF
		END_IF
		
		IF fbSeq.bError THEN
			RaiseAlarm(Id := E_Alarm.NcFeedTableRunInit, Info := fbSeq.nErrorId);
			state := E_CycleState.Abort;
		END_IF

	(*********************** End of piece, EJECT NO 2 START: wait for start **********************)
	E_CycleState.WaitStartNextPiece:
		// Pezzo finito in ciclo continuo: lo start fa il riposizionamento (50 -> 122), un altro start il pezzo.
		// Contapezzi e lotto sono gia' stati valutati nello stato 410, una volta sola.
		// Uno stop qui si applica al giro dopo; lo start della ripresa vale come questo start.
		IF stopPending THEN
			lastState := E_CycleState.CenteringSelect;
			state := E_CycleState.Stop;
		ELSIF startCondition THEN
			state := E_CycleState.CenteringSelect;
		END_IF

	(*********************** End **********************)
	E_CycleState.CycleEnd:
		//IO.clampClosedReset := TRUE;
		//IO.clampClosedSet	:= FALSE;
		state := E_CycleState.Idle;
		
	(*********************** Abort **********************)  
	E_CycleState.Abort:
		homingDone := FALSE;
		stopPending := FALSE;
		cycleEndReason := E_CycleEndReason.Aborted;

		// Arresto dei canali NC (fbNc, comando EStop dato in testa): ora si aspetta davvero la fine
		// (prima il passo leggeva bBusy del ciclo precedente e passava a 610 subito).
		IF fbNc.bDone THEN
			state := E_CycleState.AbortDone;
		END_IF

		IF fbNc.bError THEN
			RaiseAlarm(Id := E_Alarm.NcAbort, Info := fbNc.nErrorId);
			state := E_CycleState.WaitReset;
		END_IF
		
	E_CycleState.AbortDone:
		RaiseAlarm(Id := E_Alarm.CycleResetRequired);
		state := E_CycleState.WaitReset;
		
	E_CycleState.WaitReset:
		IF hmiReset THEN
			state := E_CycleState.Reset;
		END_IF
		
		IF stTwoHandControl.xStopButtonDelayTrigger THEN
			IO.clampClosedReset := TRUE;
			IO.clampClosedSet 	:= FALSE;
		END_IF
		
	(*********************** Stop **********************)  
	E_CycleState.Stop:
		// homingDone resta com'e': la ripresa da 50 o 110 deve sapere se il posizionamento iniziale e' fatto.
		// Lo azzera il Reset (800), che obbliga a rifare il posizionamento.
		stopPending := FALSE;
		cycleEndReason := E_CycleEndReason.Stopped;
		clampClosedAtStop := IO.clampClosedSet;

		// Arresto dei canali NC (fbNc, comando EStop dato in testa).
		IF fbNc.bDone THEN
			state := E_CycleState.Stopped;
		END_IF

		IF fbNc.bError THEN
			RaiseAlarm(Id := E_Alarm.NcStop, Info := fbNc.nErrorId);
			state := E_CycleState.WaitReset;
		END_IF
		
	E_CycleState.Stopped:
		IF hmiReset THEN
			state := E_CycleState.Reset;
		END_IF
		
		IF stTwoHandControl.xStopButtonDelayTrigger THEN
			IO.clampClosedReset := TRUE;
			IO.clampClosedSet 	:= FALSE;
		END_IF
		
		IF startCondition THEN
			// La morsa torna come era allo stop (lo stop tenuto premuto puo' averla aperta).
			// Dopo il posizionamento iniziale e' aperta e deve restarlo per il centraggio.
			IO.clampClosedReset := NOT clampClosedAtStop;
			IO.clampClosedSet 	:= clampClosedAtStop;
			state := E_CycleState.Resume;
		END_IF

	(*********************** Resume after stop **********************)
	// lastState = E_CycleState.SeqRun (RUN): step-on NC, i canali riprendono dal punto di arresto.
	// Altrimenti (cambio sequenza, fine centraggio, fine posizionamento iniziale, attesa start): reset dei
	// canali e ripartenza dallo stato memorizzato; il cambio sequenza riparte da 120 con lo stesso seqIdx.
	E_CycleState.Resume:
		IF lastState = E_CycleState.SeqRun THEN
			// Step-on dei canali NC (fbNc, comando StepOn dato in testa).
			IF fbNc.bDone THEN
				state := E_CycleState.SeqRun;
			END_IF

			IF fbNc.bError THEN
				RaiseAlarm(Id := E_Alarm.NcStepOn, Info := fbNc.nErrorId);
				state := E_CycleState.WaitReset;
			END_IF
		ELSE
			state := E_CycleState.ResumeResetTables;
		END_IF

	E_CycleState.ResumeResetTables:
		// Reset delle tabelle e dei canali NC nel runner (comando ResetTables, anche a meta' invio):
		// primo giro qui, la fine si legge nel passo 745.
		state := E_CycleState.ResumeResetWait;

	E_CycleState.ResumeResetWait:
		IF fbSeq.bResetDone THEN
			FOR i:=0 TO 2 DO
				channelDone[i] := FALSE;
				syncAck[i] := FALSE;
			END_FOR

			// Sincronismi della sequenza interrotta: si riparte puliti, come dallo stato 110.
			USELDone := FALSE;
			USERDone := FALSE;
			UR2Done	:= FALSE;
			USEL_UR2_Ack := FALSE;
			USER_UR2_Ack := FALSE;
			UR2_USEL_Req := FALSE;
			UR2_USER_Req := FALSE;

			// lastState = SeqPrepare (cambio sequenza): si rifa' la preparazione della sequenza corrente, seqIdx invariato.
			state := lastState;
		END_IF

		IF fbSeq.bError THEN
			RaiseAlarm(Id := E_Alarm.NcResumeReset, Info := fbSeq.nErrorId);
			state := E_CycleState.WaitReset;
		END_IF

	(*********************** Reset **********************)  
	E_CycleState.Reset:
		ClearAlarms();
		startCondition  := FALSE;   //
		stopPending := FALSE;
		// Dopo un Reset il pezzo in macchina non e' piu' seguito: il prossimo start rifa' il posizionamento iniziale.
		homingDone := FALSE;
		// Reset MC degli assi in uso (FB_AxisModule, action AxisModules): esito dal ciclo precedente.
		resetAxesCmd := TRUE;

		IF axesResetDone THEN
			state := E_CycleState.Idle;
		END_IF

		IF axesResetError THEN
			RaiseAlarm(Id := E_Alarm.NcResetAxes, Info := axesResetErrorId);
			state := E_CycleState.WaitReset;
		END_IF
		
	E_CycleState.ResetChannels:
		// Reset dei canali NC (fbNc, comando Reset dato in testa).
		IF fbNc.bDone THEN
			state := E_CycleState.Idle;
		END_IF

		IF fbNc.bError THEN
			// stato non raggiunto da nessuna transizione: nessun allarme dedicato
			state := E_CycleState.WaitReset;
		END_IF

	(*********************** New program loaded from the HMI **********************)
	E_CycleState.NewProgram:
		// Reset del ciclo dopo il caricamento di un nuovo programma dall'HMI.
		newProgramPending := FALSE;

		count := 0;
		seqIdx := 0;

		// forza la sequenza di INIT con i dati del nuovo programma
		homingDone := FALSE;

		USELDone := FALSE;
		USERDone := FALSE;
		UR2Done	:= FALSE;
		USEL_UR2_Ack := FALSE;
		USER_UR2_Ack := FALSE;
		UR2_USEL_Req := FALSE;
		UR2_USER_Req := FALSE;

		FOR i:=0 TO 2 DO
			channelDone[i] := FALSE;
			syncAck[i] := FALSE;
		END_FOR

		startCondition := FALSE;

		// il reset standard azzera la lista messaggi e riabilita gli assi
		state := E_CycleState.Reset;


	(*********************** Switch to Manual Mode **********************)
	E_CycleState.ToManual:
		homingDone := FALSE;
		stopPending := FALSE;
		cycleEndReason := E_CycleEndReason.ManualMode;

		IF udiItpState[0] > 2 AND  udiItpState[1] > 2 AND udiItpState[2] > 2 THEN
			state := E_CycleState.ToManualEStop;
		ELSE
			state := E_CycleState.ToManualClearGroups;
		END_IF
		
	E_CycleState.ToManualEStop:
		// Arresto dei canali NC (fbNc, comando EStop dato in testa).
		IF fbNc.bDone THEN
			state := E_CycleState.ToManualClearGroups;
		END_IF

		IF fbNc.bError THEN
			RaiseAlarm(Id := E_Alarm.NcManualEStop, Info := fbNc.nErrorId);
			state := E_CycleState.WaitReset;
		END_IF
		
	E_CycleState.ToManualClearGroups:
		FOR i:=0 TO 2 DO
			fbClearGroup[i](
				nGroupId:=i+7,
				bExecute:=TRUE,
				tTimeOut:=T#100MS );
		END_FOR
		
		IF (NOT fbClearGroup[0].bBusy) AND (NOT fbClearGroup[1].bBusy) AND (NOT fbClearGroup[2].bBusy) THEN
			fbClearGroup[0]( bExecute:=FALSE );
			fbClearGroup[1]( bExecute:=FALSE );
			fbClearGroup[2]( bExecute:=FALSE );
			state := E_CycleState.ToManualCheckAxes;
		END_IF
		
		IF fbClearGroup[0].bErr OR fbClearGroup[1].bErr OR fbClearGroup[2].bErr THEN
			RaiseAlarm(Id := E_Alarm.NcManualClearGroup, Info := MAX(fbClearGroup[0].nErrId, fbClearGroup[1].nErrId, fbClearGroup[2].nErrId));
			state := E_CycleState.WaitReset;
		END_IF
		
	E_CycleState.ToManualCheckAxes:
		IF ERL.Status.Error OR ERR.Status.Error OR USEL.Status.Error OR USER.Status.Error OR UR2.Status.Error THEN
			state := E_CycleState.ToManualResetAxes;
		ELSE
			state := E_CycleState.Manual;
		END_IF
	
	E_CycleState.ToManualResetAxes:
		// Reset MC degli assi in uso (FB_AxisModule, action AxisModules): esito dal ciclo precedente.
		resetAxesCmd := TRUE;

		IF axesResetDone THEN
			state := E_CycleState.Manual;
		END_IF

		IF axesResetError THEN
			RaiseAlarm(Id := E_Alarm.NcManualResetAxes, Info := axesResetErrorId);
			state := E_CycleState.WaitReset;
		END_IF
		
		
	(*********************** Manual Mode **********************) 
	E_CycleState.Manual:
		autoMode := FALSE;
		manualMode := TRUE;		
		state := E_CycleState.Idle;

		
	(*********************** Switch to Auto Mode **********************) 
	E_CycleState.ToAuto:
		autoMode := TRUE;
		manualMode := FALSE;
		state := E_CycleState.Idle;
END_CASE


//*******************************************************************************************************************
// New program loaded from the HMI
//*******************************************************************************************************************
IF newProgramTrigger THEN
	newProgramPending := TRUE;
END_IF

// Il reset ciclo viene applicato solo a programma fermo. Se la macchina sta eseguendo,
// lo stato 410 chiude il ciclo corrente e poi si passa da qui.
// Valutato prima dei Forced States, per non coprire uno stop o un abort forzato nello stesso ciclo.
IF newProgramPending AND (state = E_CycleState.Idle OR state >= E_CycleState.Abort) AND state <> E_CycleState.Reset AND state <> E_CycleState.ResetChannels THEN
	state := E_CycleState.NewProgram;
END_IF

//*******************************************************************************************************************
// Forced States
//*******************************************************************************************************************
IF state <> E_CycleState.Idle AND state < E_CycleState.Abort THEN
	// Stop. In RUN e nel cambio sequenza la macchina si ferma subito (700) e la ripresa parte da lastState.
	// Durante centraggio (55-90), posizionamento iniziale (122-412) e attesa start di fine pezzo (420) lo stop
	// si memorizza: la fase finisce e la macchina si ferma alla fine (stati 80, 90, 412, 420).
	// Le corse PTP del centraggio non si fermano comunque con lo stop (scelta confermata).
	IF hmiStop OR stTwoHandControl.xStopRTrigger THEN
		CASE state OF
			E_CycleState.Centering,
			E_CycleState.HomingPrepare, E_CycleState.HomingRun, E_CycleState.WaitStartNextPiece:
				stopPending := TRUE;
		ELSE
			lastState := state;
			state := E_CycleState.Stop;
		END_CASE
	END_IF
	
	IF NOT allDrivesEnabled THEN
		state := E_CycleState.Abort;
	END_IF
	
	IF drivesError THEN
		state := E_CycleState.Abort;
	END_IF
	
	IF NOT Safety.AbilitazionePeriferiche THEN
		//state := E_CycleState.Abort;
	END_IF
ELSE
	IF hmiProgramLoadedCmd THEN
		count := 0;
	END_IF
END_IF

IF state < E_CycleState.Abort OR (state >= E_CycleState.Stop AND state < E_CycleState.Reset) THEN
	//if manual mode is selected switch to manual mode
	IF manualModeTrigger THEN
		state := E_CycleState.ToManual;
	END_IF
END_IF

IF (state >= E_CycleState.Manual AND state < E_CycleState.ToAuto) OR state = E_CycleState.Idle THEN
	IF autoModeTrigger THEN
		state := E_CycleState.ToAuto;
	END_IF
END_IF

//*******************************************************************************************************************
// Watchdog dei passi tecnici
//*******************************************************************************************************************
// I passi che aspettano solo un FB NC/MC (reset e costruzione gruppi, tabelle, e-stop, step-on, reset assi)
// durano pochi cicli. Se uno resta fermo oltre tStateTimeOut la macchina va in abort con il passo nell'Info,
// invece di restare ferma senza messaggio. Le attese dell'operatore (0, 412, 420, 620, 719) e il RUN non sono controllati.
IF state <> stateWatchPrev THEN
	stateWatchPrev := state;
	fbStateWatchdog(IN := FALSE);
END_IF

CASE state OF
	E_CycleState.SeqPrepare, E_CycleState.HomingPrepare,
	E_CycleState.Abort, E_CycleState.Stop, E_CycleState.Resume, E_CycleState.ResumeResetTables, E_CycleState.ResumeResetWait,
	E_CycleState.Reset, E_CycleState.ResetChannels,
	E_CycleState.ToManualEStop, E_CycleState.ToManualClearGroups, E_CycleState.ToManualResetAxes:
		stateIsTechnical := TRUE;
ELSE
	stateIsTechnical := FALSE;
END_CASE

fbStateWatchdog(IN := stateIsTechnical, PT := tStateTimeOut);

IF fbStateWatchdog.Q THEN
	RaiseAlarm(Id := E_Alarm.StateTimeout, Info := state);
	fbStateWatchdog(IN := FALSE);
	IF state < E_CycleState.Abort THEN
		state := E_CycleState.Abort;
	ELSE
		state := E_CycleState.WaitReset;
	END_IF
END_IF

//*******************************************************************************************************************
// State Machine Info
//*******************************************************************************************************************
programIdle := state = E_CycleState.Idle;
programCanExecute := NOT drivesError AND allDrivesEnabled AND ProgramDB.sequence[0].active AND autoMode
	AND NOT calibrationBusy;
programAborted := state >= E_CycleState.Abort AND state <= E_CycleState.WaitReset;
programStopped := state >= E_CycleState.Stop AND state <= E_CycleState.ResumeResetWait;
programRunning := state <> E_CycleState.Idle AND state < E_CycleState.Abort;

IO.centeringLeftReset := io.centringSet;
END_ACTION

END_PROGRAM

// ---- POUs/MPG/MPG_ReadStatus.TcPOU
{attribute 'hide_all_locals'}
FUNCTION_BLOCK MPG_ReadStatus
VAR_INPUT
	uismoothingPercentage			: UINT;
	tUpdateTimerPt					: TIME;
	uiScalingFactorNumerator		: UINT;
	uiScalingFactorDenominator		: UINT;
END_VAR

VAR_IN_OUT
	stMpgEncoder 					: ST_MpgEncoder;
END_VAR

VAR
	fbUpdateTimer					: TON;
	fbButton1RTrigger				: R_TRIG;
	fbButton2RTrigger				: R_TRIG;
	fbButton3RTrigger				: R_TRIG;
	fbFowardRTrigger				: R_TRIG;
	fbBackwardRTrigger				: R_TRIG;
	fbSafetySwitchRTrigger			: R_TRIG;
	fbButton1FTrigger				: F_TRIG;
	fbButton2FTrigger				: F_TRIG;
	fbButton3FTrigger				: F_TRIG;
	fbFowardFTrigger				: F_TRIG;
	fbBackwardFTrigger				: F_TRIG;
	fbSafetySwitchFTrigger			: F_TRIG;
	_xUpdateTimerStart				: BOOL;
	_xUpdateTimerOut				: BOOL;
	_xButton1TriggerClk				: BOOL;
	_xButton2TriggerClk				: BOOL;
	_xButton3TriggerClk				: BOOL;
	_xForwardTriggerClk				: BOOL;
	_xBackwardTriggerClk			: BOOL;
	_xSafetySwitchTriggerClk		: BOOL;
	_xButton1TriggerRising			: BOOL;
	_xButton2TriggerRising			: BOOL;
	_xButton3TriggerRising 			: BOOL;
	_xForwardTriggerRising			: BOOL;
	_xBackwardTriggerRising			: BOOL;
	_xSafetySwtichTriggerRising		: BOOL;
	_xButton1TriggerFalling			: BOOL;
	_xButton2TriggerFalling			: BOOL;
	_xButton3TriggerFalling 		: BOOL;
	_xForwardTriggerFalling			: BOOL;
	_xBackwardTriggerFalling		: BOOL;
	_xSafetySwtichTriggerFalling	: BOOL;
	_uiState						: UINT;
	_rUpdateStartPosition			: REAL;
	_rUpdateEndPosition				: REAL;
	_rRawPosition					: REAL;
	_rActPosition					: REAL;
	_rSpeedAct						: REAL;
	_uiIndex						: UINT;
	_uiReadsCount					: UINT;
	_uiSum							: REAL;
	_aReadings						: ARRAY[0..200] OF REAL;
	_uiReadingsCount				: UINT;
	_rAverage						: REAL;
	_eDirection						: MC_Direction;
	_iDirection						: INT;
	_uiOverrideSpeed				: UINT;
	_uiSpeedDivider					: UINT;
	_diSelector2					: UINT;
END_VAR

//*******************************************************************************************************************
// Mapping inputs 
//*******************************************************************************************************************
_rRawPosition				:= DINT_TO_REAL(stMpgEncoder.diRowPositionFeedBack);
_rActPosition 				:= (_rRawPosition * uiScalingFactorNumerator) / uiScalingFactorDenominator;
_uiReadsCount 				:= (SIZEOF(_aReadings)/SIZEOF(REAL)) - (100 - uismoothingPercentage);
_xButton1TriggerClk			:= stMpgEncoder.diButton1;
_xButton2TriggerClk			:= stMpgEncoder.diButton2;
_xButton3TriggerClk			:= stMpgEncoder.diButton3;
_diSelector2				:= stMpgEncoder.diSelector2; 

//The selectors 1 and 2 uses a Gray-code encoder selector
//stMpgEncoder.diSelector1.2 := stMpgEncoder.diSelector1Bit3;
//stMpgEncoder.diSelector1.1 := stMpgEncoder.diSelector1.2 XOR stMpgEncoder.diSelector1Bit2;
//stMpgEncoder.diSelector1.1 := stMpgEncoder.diSelector1.1 XOR stMpgEncoder.diSelector1Bit1;
// Selettore 1 con codifica binaria
stMpgEncoder.diSelector1.2 := stMpgEncoder.diSelector1Bit3;
stMpgEncoder.diSelector1.1 := stMpgEncoder.diSelector1Bit2;
stMpgEncoder.diSelector1.0 := stMpgEncoder.diSelector1Bit1;

stMpgEncoder.diSelector2.1 := stMpgEncoder.diSelector2Bit2;
stMpgEncoder.diSelector2.0 := stMpgEncoder.diSelector2Bit1;
_xSafetySwitchTriggerClk    := stMpgEncoder.diSafetySwitch;

//*******************************************************************************************************************
// State machine
//*******************************************************************************************************************
CASE _uiState OF
	0:
		_rUpdateStartPosition 	:= _rActPosition;
		_xUpdateTimerStart 		:= TRUE;
		_uiState				:= 10;
	
	10:
		IF _xUpdateTimerOut THEN
			_xUpdateTimerStart 		:= FALSE;
			_rUpdateEndPosition 	:= _rActPosition;
			_rSpeedAct 				:= (_rUpdateEndPosition - _rUpdateStartPosition) / TIME_TO_REAL(fbUpdateTimer.ET);
			_uiSum 					:= _uiSum - _aReadings[_uiIndex];
			_aReadings[_uiIndex] 	:= _rSpeedAct;
			_uiSum 					:= _uiSum + _aReadings[_uiIndex];
			_uiIndex 				:= _uiIndex + 1;
			
			IF (_uiIndex >= _uiReadsCount) THEN
				_uiIndex := 0;
			END_IF
			
			_rAverage 				:= _uiSum / _uiReadsCount;
			_uiState				:= 0;
		END_IF
END_CASE

IF ABS(_rSpeedAct) > 0.1 THEN
	_uiOverrideSpeed 	:= REAL_TO_UINT((ABS(_rAverage) * 100) / stMpgEncoder.uiMaxSpeed);
	_iDirection 		:= REAL_TO_INT(_rAverage / ABS(_rAverage));
ELSE
	_uiOverrideSpeed := 0;
	_iDirection := 0;
END_IF

CASE _iDirection OF
	0:
		_eDirection := MC_Direction.MC_Shortest_Way;
	1:
		_eDirection := MC_Direction.MC_Positive_Direction;
	-1:
		_eDirection := MC_Direction.MC_Negative_Direction;
END_CASE

_xForwardTriggerClk := _eDirection = MC_Direction.MC_Positive_Direction;
_xBackwardTriggerClk := _eDirection = MC_Direction.MC_Negative_Direction;

CASE _diSelector2 OF
	1:
		_uiSpeedDivider := 10;
	2:
		_uiSpeedDivider := 20;
	3:
		_uiSpeedDivider := 50;
END_CASE

//*******************************************************************************************************************
// FB calls
//*******************************************************************************************************************
fbUpdateTimer(in := _xUpdateTimerStart, PT := tUpdateTimerPt, Q => _xUpdateTimerOut);
fbButton1RTrigger(Q => _xButton1TriggerRising, CLK := _xButton1TriggerClk);
fbButton2RTrigger(Q => _xButton2TriggerRising, CLK := _xButton2TriggerClk);
fbButton3RTrigger(Q => _xButton3TriggerRising, CLK := _xButton3TriggerClk);
fbFowardRTrigger(Q => _xForwardTriggerRising, CLK := _xForwardTriggerClk);
fbBackwardRTrigger(Q => _xBackwardTriggerRising, CLK := _xBackwardTriggerClk);
fbSafetySwitchRTrigger(Q => _xSafetySwtichTriggerRising, CLK := _xSafetySwitchTriggerClk);
fbButton1FTrigger(Q => _xButton1TriggerFalling, CLK := _xButton1TriggerClk);
fbButton2FTrigger(Q => _xButton2TriggerFalling, CLK := _xButton2TriggerClk);
fbButton3FTrigger(Q => _xButton3TriggerFalling, CLK := _xButton3TriggerClk);
fbFowardFTrigger(Q => _xForwardTriggerFalling, CLK := _xForwardTriggerClk);
fbBackwardFTrigger(Q => _xBackwardTriggerFalling, CLK := _xBackwardTriggerClk);
fbSafetySwitchFTrigger(Q => _xSafetySwtichTriggerFalling, CLK := _xSafetySwitchTriggerClk);



//*******************************************************************************************************************
// Mapping  outputs  
//*******************************************************************************************************************
stMpgEncoder.rActPos 			:= _rActPosition;
stMpgEncoder.rActVelo			:= _rAverage;
stMpgEncoder.eDirection 		:= _eDirection;
stMpgEncoder.uiOverrideSpeed	:= _uiOverrideSpeed;
stMpgEncoder.xButton1RTrigger	:= _xButton1TriggerRising;
stMpgEncoder.xButton2RTrigger	:= _xButton2TriggerRising;
stMpgEncoder.xButton3RTrigger	:= _xButton3TriggerRising;
stMpgEncoder.xFowardRTrigger		:= _xForwardTriggerRising;
stMpgEncoder.xBackwardRTrigger	:= _xBackwardTriggerRising;
stMpgEncoder.uiSpeedDivider		:= _uiSpeedDivider;
stMpgEncoder.xSafetySwitchRTrigger := _xSafetySwtichTriggerRising;
stMpgEncoder.xButton1FTrigger	:= _xButton1TriggerFalling;
stMpgEncoder.xButton2FTrigger	:= _xButton2TriggerFalling;
stMpgEncoder.xButton3FTrigger	:= _xButton3TriggerFalling;
stMpgEncoder.xFowardFTrigger		:= _xForwardTriggerFalling;
stMpgEncoder.xBackwardFTrigger	:= _xBackwardTriggerFalling;
stMpgEncoder.xSafetySwitchFTrigger := _xSafetySwtichTriggerFalling;

END_FUNCTION_BLOCK

// ---- POUs/TwoHand/TwoHand_ReadStatus.TcPOU
{attribute 'hide_all_locals'}
FUNCTION_BLOCK TwoHand_ReadStatus

VAR_IN_OUT
	stTwoHandControl	: ST_TwoHandControl;
END_VAR

VAR
	fbButton1RTrigger				: R_TRIG;
	fbStartRTrigger					: R_TRIG;
	fbStop1RTrigger					: R_TRIG;
	fbTwoHandRTrigger				: R_TRIG;
	fbSafetySwitchRTrigger			: R_TRIG;
	fbStopButtonDelayTrigger		: R_TRIG;
	fbButton1FTrigger				: F_TRIG;
	fbStartFTrigger					: F_TRIG;
	fbStop1FTrigger					: F_TRIG;
	fbTwoHandFTrigger				: F_TRIG;
	fbSafetySwitchFTrigger			: F_TRIG;
	fbStopButtonTimer				: TON;
	_xButton1TriggerClk				: BOOL;
	_xStartTriggerClk				: BOOL;
	_xStopTriggerClk				: BOOL;
	_XStopButtonDelayClk			: BOOL;
	_xTwoHandTriggerClk				: BOOL;
	_xSafetySwitchTriggerClk		: BOOL;
	_xButton1TriggerRising			: BOOL;
	_xStartTriggerRising			: BOOL;
	_xStopTriggerRising				: BOOL;
	_xTwoHandTriggerRising			: BOOL;
	_xSafetySwitchTriggerRising		: BOOL;
	_xButton1TriggerFalling			: BOOL;
	_xStartTriggerFalling			: BOOL;
	_xStopTriggerFalling			: BOOL;
	_xTwoHandTriggerFalling			: BOOL;
	_xSafetySwitchTriggerFalling	: BOOL;
	_xStopButtonDelayRising			: BOOL;
END_VAR

//*******************************************************************************************************************
// Mapping inputs 
//*******************************************************************************************************************
_xButton1TriggerClk			:= stTwoHandControl.diButton1;	
_xStartTriggerClk			:= stTwoHandControl.diStartButton;		
_xStopTriggerClk			:= stTwoHandControl.diStopButton;		
_xTwoHandTriggerClk			:= stTwoHandControl.diTwoHand;		
_xSafetySwitchTriggerClk	:= stTwoHandControl.diSafetySwitch;		

//*******************************************************************************************************************
// FB calls
//*******************************************************************************************************************
fbButton1RTrigger(CLK := _xButton1TriggerClk, Q => _xButton1TriggerRising);
fbStartRTrigger(CLK := _xStartTriggerClk, Q => _xStartTriggerRising);
fbStop1RTrigger(CLK := _xStopTriggerClk, Q => _xStopTriggerRising);
fbTwoHandRTrigger(CLK := _xTwoHandTriggerClk, Q => _xTwoHandTriggerRising);
fbSafetySwitchRTrigger(CLK := _xSafetySwitchTriggerClk, Q => _xSafetySwitchTriggerRising);

fbButton1FTrigger(CLK := _xButton1TriggerClk, Q => _xButton1TriggerFalling);
fbStartFTrigger(CLK := _xStartTriggerClk, Q => _xStartTriggerFalling);
fbStop1FTrigger(CLK := _xStopTriggerClk, Q => _xStopTriggerFalling);
fbTwoHandFTrigger(CLK := _xTwoHandTriggerClk, Q => _xTwoHandTriggerFalling);
fbSafetySwitchFTrigger(CLK := _xSafetySwitchTriggerClk, Q => _xSafetySwitchTriggerFalling);

fbStopButtonTimer(IN := _xStopTriggerClk, PT := T#1000MS, Q => _xStopButtonDelayClk);

fbStopButtonDelayTrigger(CLK := _xStopButtonDelayClk, Q =>_xStopButtonDelayRising);
//*******************************************************************************************************************
// Mapping  outputs  
//*******************************************************************************************************************
stTwoHandControl.xButton1RTrigger		:= _xButton1TriggerRising;
stTwoHandControl.xStartRTrigger			:= _xStartTriggerRising;
stTwoHandControl.xStopRTrigger			:= _xStopTriggerRising;
stTwoHandControl.xTwoHandRTrigger		:= _xTwoHandTriggerRising;
stTwoHandControl.xSafetySwitchRTrigger	:= _xSafetySwitchTriggerRising;

stTwoHandControl.xButton1FTrigger		:= _xButton1TriggerFalling;
stTwoHandControl.xStartFTrigger			:= _xStartTriggerFalling;
stTwoHandControl.xStopFTrigger			:= _xStopTriggerFalling;
stTwoHandControl.xTwoHandFTRigger		:= _xTwoHandTriggerFalling;
stTwoHandControl.xSafetySwitchFTrigger	:= _xSafetySwitchTriggerFalling;
stTwoHandControl.xStopButtonDelayTrigger := _xStopButtonDelayRising;

END_FUNCTION_BLOCK

// ---- Core/Nc/FB_SequenceRunner.TcPOU
// Le tabelle NC di una sequenza di ProgramDB, per tutti i canali: preparazione, esecuzione, reset.
// La stessa per le sequenze del pezzo e per l'homing (prima erano due catene di passi uguali, 120-402).
// Va chiamato a ogni ciclo PLC con il comando del ciclo (eCmd):
// - Prepare: reset gruppi -> costruzione gruppi -> reset tabelle -> GeoStart -> riempimento -> invio; poi bReady;
// - Run: legge la fine dei canali (aChannelDone, non memorizzata: la memorizza il ciclo);
// - ResetTables: reset di FB_NciFeedTable (tabella interrotta e canale NC dopo un arresto); poi bResetDone;
// - None: solo i FB dei gruppi, che devono girare sempre.
// Un comando diverso dal ciclo precedente riparte da capo. Gli errori restano in bError (con il passo e
// l'ErrorID) finche' il comando non cambia: l'allarme lo sceglie il ciclo.
FUNCTION_BLOCK FB_SequenceRunner
VAR_INPUT
	eCmd					: E_SeqCmd;
	pSequence				: POINTER TO TYPE_SEQUENCE;	// sequenza da preparare/eseguire (homing o ProgramDB.sequence[i])
	nGroupIdBase			: UDINT := 7;		// ID NC del gruppo del canale 0
	tGroupTimeOut			: TIME := T#100MS;	// timeout dei comandi ai gruppi
	bCenteringCorrection	: BOOL;				// centraggio TB: correzione delle quote
	fToleranceMeasure		: LREAL;			// tolleranza misurata dal centraggio
	bSingleBlock			: BOOL;				// passo-passo: le M di start entrano in tabella
	nDefCount				: UINT;				// righe valide di aDef
	bLogFeederEntries		: BOOL;				// log delle righe inviate (FB_NciFeedTable)
END_VAR
VAR_IN_OUT
	aNciToPlc				: ARRAY[0..Core_Param.MAX_CHANNEL-1] OF NCTOPLC_NCICHANNEL_REF;
	aAxisCfg				: ARRAY[*] OF ST_AxisCfg;
	aDef					: ARRAY[*] OF ST_MFuncDef;
END_VAR
VAR_OUTPUT
	eStep					: E_SeqStep;
	bReady					: BOOL;		// Prepare: tabelle inviate ai canali
	bResetDone				: BOOL;		// ResetTables: reset finito
	aChannelDone			: ARRAY[0..Core_Param.MAX_CHANNEL-1] OF BOOL;	// Run: il canale ha finito (bChannelDone)
	bError					: BOOL;
	eErrorStep				: E_SeqStep;	// passo in cui e' nato l'errore
	nErrorId				: UDINT;		// ErrorID del FB NC (0 se non c'e')
END_VAR
VAR
	eLastCmd				: E_SeqCmd;
	fbClearGroups			: FB_ClearInterpolationGroup;
	fbBuildGroups			: FB_BuildGroups;
	fbTablePrep				: ARRAY[0..Core_Param.MAX_CHANNEL-1] OF FB_NciFeedTablePreparation;
	fbBuilder				: FB_FeedTableBuilder;
	fbFeedTable				: ARRAY[0..Core_Param.MAX_CHANNEL-1] OF FB_NciFeedTable;
	aFeedGroupTable			: ARRAY[0..Core_Param.MAX_CHANNEL-1] OF ST_NciFeedGroupTable;
	stGeoStart				: ARRAY[0..Core_Param.MAX_CHANNEL-1] OF ST_NciGeoStart;
	bClearExecute			: BOOL;
	bBuildExecute			: BOOL;
	nResetScans				: UINT;
	bAnyBusy				: BOOL;
	ch						: UINT;
	i						: UINT;
	nAxis					: UINT;
END_VAR

bClearExecute := FALSE;
bBuildExecute := FALSE;
bReady := FALSE;
bResetDone := FALSE;

IF eCmd <> eLastCmd THEN
	eLastCmd := eCmd;
	bError := FALSE;
	eErrorStep := E_SeqStep.Idle;
	nErrorId := 0;
	CASE eCmd OF
		E_SeqCmd.Prepare:		eStep := E_SeqStep.ClearGroups;
		E_SeqCmd.Run:			eStep := E_SeqStep.Running;
		E_SeqCmd.ResetTables:	eStep := E_SeqStep.Resetting;
								nResetScans := 0;
	ELSE
		eStep := E_SeqStep.Idle;
	END_CASE
END_IF

IF eStep >= E_SeqStep.ClearGroups AND eStep <= E_SeqStep.Running AND pSequence = 0 THEN
	Fail(eStep, 0);
END_IF

CASE eStep OF
	E_SeqStep.ClearGroups:
		// I FB dei gruppi girano in fondo: qui si legge l'esito della chiamata precedente.
		bClearExecute := TRUE;
		IF fbClearGroups.bDone THEN
			eStep := E_SeqStep.BuildGroups;
		END_IF
		IF fbClearGroups.bError THEN
			Fail(E_SeqStep.ClearGroups, 0);
		END_IF

	E_SeqStep.BuildGroups:
		bBuildExecute := TRUE;
		IF fbBuildGroups.bDone THEN
			eStep := E_SeqStep.TableReset;
		END_IF
		IF fbBuildGroups.bError THEN
			Fail(E_SeqStep.BuildGroups, 0);
		END_IF

	E_SeqStep.TableReset:
		FOR ch := 0 TO Core_Param.MAX_CHANNEL - 1 DO
			IF pSequence^.task[ch].active THEN
				fbTablePrep[ch](bResetAll := TRUE, stFeedGroupTable := aFeedGroupTable[ch]);
			END_IF
			fbTablePrep[ch].bResetAll := FALSE;
		END_FOR
		CheckTablePrep(E_SeqStep.TableReset);
		IF NOT bError THEN
			eStep := E_SeqStep.TableStart;
		END_IF

	E_SeqStep.TableStart:
		// Punto di partenza = posizione attuale degli assi del gruppo, nell'ordine di FB_BuildGroups (X, Y, Z).
		// FB_FeedTableBuilder poi azzera la tabella (come faceva FB_FeedTablesPrep): il passo resta per fedelta'.
		FOR ch := 0 TO Core_Param.MAX_CHANNEL - 1 DO
			IF pSequence^.task[ch].active THEN
				FOR i := 0 TO 2 DO
					nAxis := TO_UINT(pSequence^.task[ch].axisGroup[i]);
					IF nAxis >= LOWER_BOUND(aAxisCfg, 1) AND nAxis <= UPPER_BOUND(aAxisCfg, 1) THEN
						CASE i OF
							0: stGeoStart[ch].fPosX := aAxisCfg[nAxis].fActPos;
							1: stGeoStart[ch].fPosY := aAxisCfg[nAxis].fActPos;
							2: stGeoStart[ch].fPosZ := aAxisCfg[nAxis].fActPos;
						END_CASE
					END_IF
				END_FOR
				fbTablePrep[ch](
					nEntryType			:= E_NciEntryTypeGeoStart,
					pEntry				:= ADR(stGeoStart[ch]),
					bResetAll			:= FALSE,
					bResetTable			:= FALSE,
					stFeedGroupTable	:= aFeedGroupTable[ch]);
			END_IF
		END_FOR
		CheckTablePrep(E_SeqStep.TableStart);
		IF NOT bError THEN
			eStep := E_SeqStep.TableFill;
		END_IF

	E_SeqStep.TableFill:
		fbBuilder(
			pSequence				:= pSequence,
			bCenteringCorrection	:= bCenteringCorrection,
			fToleranceMeasure		:= fToleranceMeasure,
			bSingleBlock			:= bSingleBlock,
			nDefCount				:= nDefCount,
			aFeedGroupTable			:= aFeedGroupTable,
			aAxisCfg				:= aAxisCfg,
			aDef					:= aDef);
		IF fbBuilder.bError THEN
			Fail(E_SeqStep.TableFill, fbBuilder.nErrorId);
		ELSE
			eStep := E_SeqStep.TableFeed;
		END_IF

	E_SeqStep.TableFeed:
		bAnyBusy := FALSE;
		FOR ch := 0 TO Core_Param.MAX_CHANNEL - 1 DO
			IF pSequence^.task[ch].active THEN
				fbFeedTable[ch](
					bExecute			:= TRUE,
					bReset				:= FALSE,
					bLogFeederEntries	:= bLogFeederEntries,
					stFeedGroupTable	:= aFeedGroupTable[ch],
					stNciToPlc			:= aNciToPlc[ch]);
				IF fbFeedTable[ch].bError AND NOT bError THEN
					Fail(E_SeqStep.TableFeed, fbFeedTable[ch].nErrorId);
				END_IF
			END_IF
			bAnyBusy := bAnyBusy OR fbFeedTable[ch].bFeedBusy;
		END_FOR

		IF NOT bAnyBusy AND NOT bError THEN
			FOR ch := 0 TO Core_Param.MAX_CHANNEL - 1 DO
				fbFeedTable[ch](bExecute := FALSE, bReset := FALSE, stFeedGroupTable := aFeedGroupTable[ch], stNciToPlc := aNciToPlc[ch]);
			END_FOR
			eStep := E_SeqStep.Ready;
			bReady := TRUE;		// gia' in questo ciclo, come prima il passaggio 400 -> 410
		END_IF

	E_SeqStep.Ready:
		bReady := TRUE;

	E_SeqStep.Running:
		FOR ch := 0 TO Core_Param.MAX_CHANNEL - 1 DO
			aChannelDone[ch] := FALSE;
			IF pSequence^.task[ch].active THEN
				fbFeedTable[ch](bExecute := FALSE, bReset := FALSE, stFeedGroupTable := aFeedGroupTable[ch], stNciToPlc := aNciToPlc[ch]);
				aChannelDone[ch] := fbFeedTable[ch].bChannelDone;
				IF fbFeedTable[ch].bError AND NOT bError THEN
					Fail(E_SeqStep.Running, fbFeedTable[ch].nErrorId);
				END_IF
			END_IF
		END_FOR

	E_SeqStep.Resetting:
		// Reset di FB_NciFeedTable su tutti i canali: azzera la tabella interrotta e resetta il canale NC
		// dopo l'arresto (ItpResetEx2 interno). bResetBusy si legge dal secondo ciclo.
		bAnyBusy := FALSE;
		FOR ch := 0 TO Core_Param.MAX_CHANNEL - 1 DO
			fbFeedTable[ch](bExecute := FALSE, bReset := TRUE, stFeedGroupTable := aFeedGroupTable[ch], stNciToPlc := aNciToPlc[ch]);
			bAnyBusy := bAnyBusy OR fbFeedTable[ch].bResetBusy;
			IF fbFeedTable[ch].bError AND NOT bError THEN
				Fail(E_SeqStep.Resetting, fbFeedTable[ch].nErrorId);
			END_IF
		END_FOR

		IF nResetScans > 0 AND NOT bAnyBusy AND NOT bError THEN
			FOR ch := 0 TO Core_Param.MAX_CHANNEL - 1 DO
				fbFeedTable[ch](bExecute := FALSE, bReset := FALSE, stFeedGroupTable := aFeedGroupTable[ch], stNciToPlc := aNciToPlc[ch]);
			END_FOR
			eStep := E_SeqStep.ResetDone;
			bResetDone := TRUE;	// gia' in questo ciclo, come prima il passo 745
		END_IF
		nResetScans := nResetScans + 1;

	E_SeqStep.ResetDone:
		bResetDone := TRUE;
END_CASE

// FB dei gruppi: a ogni ciclo, come prima in MAIN.AxisFunctionBlocks; partono sul fronte di bExecute.
fbClearGroups(bExecute := bClearExecute, tTimeOut := tGroupTimeOut, nGroupIdBase := nGroupIdBase);
fbBuildGroups(bExecute := bBuildExecute, sequence := pSequence, nGroupIdBase := nGroupIdBase, aAxisCfg := aAxisCfg);

// Ferma la preparazione/esecuzione con un errore (il primo vince).
METHOD PRIVATE Fail
VAR_INPUT
	eAt			: E_SeqStep;
	nId			: UDINT;
END_VAR
IF NOT bError THEN
	bError := TRUE;
	eErrorStep := eAt;
	nErrorId := nId;
END_IF
eStep := E_SeqStep.Error;
END_METHOD

// Errore di uno dei FB_NciFeedTablePreparation dopo un passo sulle tabelle.
METHOD PRIVATE CheckTablePrep
VAR_INPUT
	eAt			: E_SeqStep;
END_VAR
VAR
	k			: UINT;
END_VAR
FOR k := 0 TO Core_Param.MAX_CHANNEL - 1 DO
	IF fbTablePrep[k].bError THEN
		Fail(eAt, fbTablePrep[k].nErrorId);
	END_IF
END_FOR
END_METHOD

END_FUNCTION_BLOCK

// ---- Core/Nc/FB_ClearInterpolationGroup.TcPOU
// Svuota i gruppi di interpolazione dei canali (ID nGroupIdBase .. nGroupIdBase + MAX_CHANNEL - 1).
{attribute 'hide_all_locals'}
FUNCTION_BLOCK FB_ClearInterpolationGroup
VAR_INPUT
	bExecute 				: BOOL;
	tTimeOut 				: TIME;
	nGroupIdBase			: UDINT := 7;	// ID NC del gruppo del canale 0
END_VAR
VAR_OUTPUT
	bDone					: BOOL;
	bBusy					: BOOL;
	bError					: BOOL;
END_VAR
VAR
	startTriggerOutput		: BOOL;
	clearGroupExecute		: BOOL;
	state					: UINT;
	groupIndex				: UINT;
	fbClearGroup			: ARRAY[0..Core_Param.MAX_CHANNEL-1] OF CfgReconfigGroup;
	fbStartTrigger			: R_TRIG;
	anyBusy					: BOOL;
	anyErr					: BOOL;
END_VAR

fbStartTrigger(CLK := bExecute, Q => startTriggerOutput);

CASE state OF
	(************************** state 0 - IDLE *************************)
	0:
		bBusy := FALSE;
		bDone := FALSE;
		clearGroupExecute := FALSE;

		IF startTriggerOutput THEN
			bBusy := TRUE;
			bError := FALSE;
			clearGroupExecute := TRUE;
			state := 10;
		END_IF

	(************** state 10 - Execute clear groups *************)
	10:
		bBusy := TRUE;

		anyBusy := FALSE;
		anyErr := FALSE;
		FOR groupIndex := 0 TO Core_Param.MAX_CHANNEL - 1 DO
			anyBusy := anyBusy OR fbClearGroup[groupIndex].bBusy;
			anyErr := anyErr OR fbClearGroup[groupIndex].bErr;
		END_FOR

		IF NOT anyBusy THEN
			state := 20;
		END_IF

		IF anyErr THEN
			state := 30;
		END_IF

	(************** state 20 - End *************)
	20:
		bDone := TRUE;
		state := 0;

	(************** state 30 - Error *************)
	30:
		bError := TRUE;
		state := 0;

END_CASE

FOR groupIndex := 0 TO Core_Param.MAX_CHANNEL - 1 DO
	fbClearGroup[groupIndex](
	nGroupId:=nGroupIdBase+groupIndex,
	bExecute:=clearGroupExecute,
	tTimeOut:=tTimeOut,
	bErr => );
END_FOR

END_FUNCTION_BLOCK

// ---- Core/Nc/FB_BuildGroups.TcPOU
// Costruisce un gruppo di interpolazione 3D per ogni task attivo della sequenza (gruppo nGroupIdBase + task):
// gli assi dell'axisGroup nell'ordine X, Y, Z, Q1, Q2. L'ID NC di ogni asse viene da aAxisCfg (indice = AXIS_ENUM).
FUNCTION_BLOCK FB_BuildGroups
VAR_INPUT
	bExecute					: BOOL;
	sequence					: POINTER TO TYPE_SEQUENCE;
	nGroupIdBase				: UDINT := 7;	// ID NC del gruppo del task 0
END_VAR
VAR_IN_OUT
	aAxisCfg					: ARRAY[*] OF ST_AxisCfg;
END_VAR
VAR_OUTPUT
	bDone						: BOOL;
	bBusy						: BOOL;
	bError						: BOOL;
END_VAR
VAR
	startTriggerOutput			: BOOL;
	buildGroupsExecute			: BOOL;
	groupCordFound				: BOOL;
	channelIndex				: UINT;
	state						: UINT;
	taskIdx						: UINT;
	AXISIdx						: UINT;
	fbStartTrigger				: R_TRIG;
	fbBuildGroup				: ARRAY[0..Core_Param.MAX_CHANNEL-1] OF CfgBuildExt3DGroup;
END_VAR

fbStartTrigger(CLK := bExecute, Q => startTriggerOutput);


CASE state OF
	(************************** state 0 - IDLE *************************)  
	0:	
		bBusy := FALSE;
		bDone := FALSE;
		buildGroupsExecute := FALSE;
		
		IF startTriggerOutput THEN
			bError := FALSE;
			state := 10;
		END_IF
		
	(************** state 10 - Prepare Groups *************)  
	10:
		bBusy := TRUE;
		taskIdx := 0;
		WHILE taskIdx < Size.MAX_TASK AND_THEN sequence^.task[taskIdx].active DO
			fbBuildGroup[taskIdx](
				nGroupId:=nGroupIdBase+taskIdx,
				nXAxisId := 0,
				nYAxisId := 0,
				nZAxisId := 0,
				nQ1AxisId := 0,
				nQ2AxisId := 0,
				nQ3AxisId := 0,
				nQ4AxisId := 0,
				nQ5AxisId := 0,
				bExecute:=FALSE );
				
			axisIdx := 0;
			
			WHILE axisIdx < Size.MAX_AXIS AND_THEN sequence^.task[taskIdx].axisGroup[axisIdx] <> AXIS_ENUM.null DO
				groupCordFound := FALSE;
				
				IF (fbBuildGroup[taskIdx].nXAxisId = 0) AND NOT groupCordFound THEN
					fbBuildGroup[taskIdx](nXAxisId := aAxisCfg[TO_UINT(sequence^.task[taskIdx].axisGroup[axisIdx])].nNcAxisId);
					groupCordFound := TRUE;
				END_IF
				
				IF (fbBuildGroup[taskIdx].nYAxisId = 0) AND NOT groupCordFound THEN
					fbBuildGroup[taskIdx](nYAxisId := aAxisCfg[TO_UINT(sequence^.task[taskIdx].axisGroup[axisIdx])].nNcAxisId);
					groupCordFound := TRUE;
				END_IF
				
				IF (fbBuildGroup[taskIdx].nZAxisId = 0) AND NOT groupCordFound THEN
					fbBuildGroup[taskIdx](nZAxisId := aAxisCfg[TO_UINT(sequence^.task[taskIdx].axisGroup[axisIdx])].nNcAxisId);
					groupCordFound := TRUE;
				END_IF
				
				IF (fbBuildGroup[taskIdx].nQ1AxisId = 0) AND NOT groupCordFound THEN
					fbBuildGroup[taskIdx](nQ1AxisId := aAxisCfg[TO_UINT(sequence^.task[taskIdx].axisGroup[axisIdx])].nNcAxisId);
					groupCordFound := TRUE;
				END_IF
				
				IF (fbBuildGroup[taskIdx].nQ2AxisId = 0) AND NOT groupCordFound THEN
					fbBuildGroup[taskIdx](nQ2AxisId := aAxisCfg[TO_UINT(sequence^.task[taskIdx].axisGroup[axisIdx])].nNcAxisId);
					groupCordFound := TRUE;
				END_IF
				
				axisIdx := axisIdx +1;
			END_WHILE
			taskIdx := taskIdx + 1;
		END_WHILE
		
		state := 20;
		
	(************** state 20 - Execute Build Group *************)  
	20:
		FOR channelIndex:=0 TO 2 DO
			fbBuildGroup[channelIndex](
			bExecute:=TRUE,
			tTimeOut:=T#100MS );
		END_FOR
		
		IF (NOT fbBuildGroup[0].bBusy) AND (NOT fbBuildGroup[1].bBusy) AND (NOT fbBuildGroup[2].bBusy) THEN
			fbBuildGroup[0]( bExecute:=FALSE );
			fbBuildGroup[1]( bExecute:=FALSE );
			fbBuildGroup[2]( bExecute:=FALSE );
			state := 100;
		END_IF
		
		IF fbBuildGroup[0].bErr OR fbBuildGroup[1].bErr OR fbBuildGroup[2].bErr THEN
			state := 200;
		END_IF
		
	(************** state 100 - End *************)  
	100:
		bDone := TRUE;
		state := 0;
		
	(************** state 200 - Error *************)  
	200:
		bError := TRUE;
		state := 0;

END_CASE

END_FUNCTION_BLOCK

// ---- Core/Nc/FB_FeedTableBuilder.TcPOU
// Riempie le tabelle NC (una per canale) con una sequenza di ProgramDB: per ogni task azzera la tabella,
// aggiunge le righe di movimento e le funzioni M nell'ordine del programma, poi la fine tabella.
// Ex FB_FeedTablesPrep, con gli assi letti dalla configurazione invece che cablati:
// - la quota di un asse va nella coordinata del gruppo NC in cui FB_BuildGroups l'ha messo
//   (1o asse dell'axisGroup = X, 2o = Y, 3o = Z), la velocita' e' speed * fSpeedScale dell'asse;
// - le funzioni M di tipo WaitStart (start del passo-passo) entrano in tabella solo con bSingleBlock.
// Si chiama una volta (un ciclo PLC) per sequenza.
FUNCTION_BLOCK FB_FeedTableBuilder
VAR_INPUT
	pSequence				: POINTER TO TYPE_SEQUENCE;
	bCenteringCorrection	: BOOL;		// centraggio TB attivo: le quote degli assi con bCenteringCorrection si correggono
	fToleranceMeasure		: LREAL;	// tolleranza misurata dal centraggio
	bSingleBlock			: BOOL;		// passo-passo: anche le funzioni M WaitStart vanno in tabella
	nDefCount				: UINT;		// righe valide di aDef
END_VAR
VAR_IN_OUT
	aFeedGroupTable			: ARRAY[0..Core_Param.MAX_CHANNEL-1] OF ST_NciFeedGroupTable;
	aAxisCfg				: ARRAY[*] OF ST_AxisCfg;
	aDef					: ARRAY[*] OF ST_MFuncDef;
END_VAR
VAR_OUTPUT
	bError					: BOOL;		// una riga non e' entrata in tabella (es. tabella piena)
	nErrorId				: UDINT;	// errore di FB_NciFeedTablePreparation
	nErrorChannel			: UINT;
END_VAR
VAR
	fbFeedTablePrep			: ARRAY[0..Core_Param.MAX_CHANNEL-1] OF FB_NciFeedTablePreparation;
	// Restano da una chiamata all'altra: una riga che non muove un asse lascia la sua ultima quota.
	stGeoLine				: ARRAY[0..Core_Param.MAX_CHANNEL-1] OF ST_NciGeoLine;
	stMFuncHsk				: ARRAY[0..Core_Param.MAX_CHANNEL-1] OF ST_NciMFuncHsk;
	stHParam				: ARRAY[0..Core_Param.MAX_CHANNEL-1] OF ST_NciHParam;
	stEndOfTables			: ARRAY[0..Core_Param.MAX_CHANNEL-1] OF ST_NciEndOfTables;
	ch						: UINT;
	actionIdx				: UINT;
	posIdx					: UINT;
	macroIdx				: UINT;
	slot					: UINT;
	nAxis					: UINT;
	fValue					: LREAL;
	bAddMacro				: BOOL;
	i						: DINT;
END_VAR

bError := FALSE;
nErrorId := 0;

// Tabelle dei task usati azzerate (come FB_FeedTablesPrep: anche il GeoStart scritto prima si perde).
FOR ch := 0 TO Core_Param.MAX_CHANNEL - 1 DO
	IF pSequence^.task[ch].active THEN
		fbFeedTablePrep[ch](bResetAll := TRUE, stFeedGroupTable := aFeedGroupTable[ch]);
		fbFeedTablePrep[ch].bResetAll := FALSE;
	END_IF
END_FOR

FOR ch := 0 TO Core_Param.MAX_CHANNEL - 1 DO
	IF pSequence^.task[ch].active THEN
		actionIdx := 0;
		WHILE actionIdx < Size.MAX_ACTION AND_THEN pSequence^.task[ch].actions[actionIdx].active DO
			CASE pSequence^.task[ch].actions[actionIdx].aType OF

				ACTION_ENUM.MOVEMENT:
					posIdx := 0;
					WHILE posIdx < Size.MAX_POSITION AND_THEN pSequence^.task[ch].actions[actionIdx].pos[posIdx].active DO
						nAxis := TO_UINT(pSequence^.task[ch].actions[actionIdx].pos[posIdx].axis);

						// Coordinata del gruppo NC in cui sta l'asse
						slot := Size.MAX_AXIS;
						FOR i := 0 TO Size.MAX_AXIS - 1 DO
							IF TO_UINT(pSequence^.task[ch].axisGroup[i]) = nAxis THEN
								slot := TO_UINT(i);
								EXIT;
							END_IF
						END_FOR

						IF (nAxis >= LOWER_BOUND(aAxisCfg, 1) AND nAxis <= UPPER_BOUND(aAxisCfg, 1))
							AND_THEN (aAxisCfg[nAxis].bDefined AND slot <= 2) THEN
							IF aAxisCfg[nAxis].bTargetZero THEN
								fValue := 0;
							ELSE
								fValue := pSequence^.task[ch].actions[actionIdx].pos[posIdx].value;
								IF aAxisCfg[nAxis].bCenteringCorrection AND bCenteringCorrection
									AND pSequence^.task[ch].actions[actionIdx].centeringVerse <> 0 THEN
									fValue := fValue + pSequence^.task[ch].actions[actionIdx].centeringAmount
										* pSequence^.task[ch].actions[actionIdx].centeringVerse * fToleranceMeasure;
								END_IF
							END_IF

							CASE slot OF
								0: stGeoLine[ch].fEndPosX := fValue;
								1: stGeoLine[ch].fEndPosY := fValue;
								2: stGeoLine[ch].fEndPosZ := fValue;
							END_CASE
							stGeoLine[ch].fVelo := pSequence^.task[ch].actions[actionIdx].speed * aAxisCfg[nAxis].fSpeedScale;
						END_IF
						posIdx := posIdx + 1;
					END_WHILE

					stGeoLine[ch].bRapidTraverse := FALSE;
					stGeoLine[ch].bAccurateStop := TRUE;
					fbFeedTablePrep[ch](
						nEntryType			:= E_NciEntryTypeGeoLine,
						pEntry				:= ADR(stGeoLine[ch]),
						bResetTable			:= FALSE,
						stFeedGroupTable	:= aFeedGroupTable[ch]);
					CheckError(ch);

				ACTION_ENUM.MACRO:
					macroIdx := 0;
					WHILE macroIdx < Size.MAX_MACRO AND_THEN pSequence^.task[ch].actions[actionIdx].macros[macroIdx].active DO
						stMFuncHsk[ch].nMFunc := UDINT_TO_INT(pSequence^.task[ch].actions[actionIdx].macros[macroIdx].mNo);
						stHParam[ch].nHParam := UDINT_TO_DINT(pSequence^.task[ch].actions[actionIdx].macros[macroIdx].delay);

						// Lo start del passo-passo serve solo in passo-passo.
						bAddMacro := TRUE;
						IF NOT bSingleBlock THEN
							i := LOWER_BOUND(aDef, 1);
							WHILE i < LOWER_BOUND(aDef, 1) + nDefCount AND_THEN i <= UPPER_BOUND(aDef, 1) DO
								IF aDef[i].nChannel = ch AND aDef[i].nMFunc = INT_TO_UINT(stMFuncHsk[ch].nMFunc) THEN
									bAddMacro := aDef[i].eKind <> E_MFuncKind.WaitStart;
									EXIT;
								END_IF
								i := i + 1;
							END_WHILE
						END_IF

						IF bAddMacro THEN
							fbFeedTablePrep[ch](
								nEntryType			:= E_NciEntryTypeHParam,
								pEntry				:= ADR(stHParam[ch]),
								bResetTable			:= FALSE,
								stFeedGroupTable	:= aFeedGroupTable[ch]);
							CheckError(ch);
							fbFeedTablePrep[ch](
								nEntryType			:= E_NciEntryTypeMFuncHsk,
								pEntry				:= ADR(stMFuncHsk[ch]),
								bResetTable			:= FALSE,
								stFeedGroupTable	:= aFeedGroupTable[ch]);
							CheckError(ch);
						END_IF
						macroIdx := macroIdx + 1;
					END_WHILE
			END_CASE
			actionIdx := actionIdx + 1;
		END_WHILE

		fbFeedTablePrep[ch](
			nEntryType			:= E_NciEntryTypeEndOfTables,
			pEntry				:= ADR(stEndOfTables[ch]),
			bResetTable			:= FALSE,
			stFeedGroupTable	:= aFeedGroupTable[ch]);
		CheckError(ch);
	END_IF
END_FOR

// Ricorda il primo errore di FB_NciFeedTablePreparation della chiamata.
METHOD PRIVATE CheckError
VAR_INPUT
	nChannel	: UINT;
END_VAR
IF fbFeedTablePrep[nChannel].bError AND NOT bError THEN
	bError := TRUE;
	nErrorId := fbFeedTablePrep[nChannel].nErrorId;
	nErrorChannel := nChannel;
END_IF
END_METHOD

END_FUNCTION_BLOCK

